(* IEC 61131-3 sources: deprecated-refusr-repo/GP/Main/samples (part 21) *)

(* ---- RND-EXPR_hewed-hoper-pudgy.st ---- *)
(*
This code implements a randomly grown symbolic expression:

((IN43 & IN39) | (!((IN20 & ((IN38 | (!(xor(xor(!(IN25), IN22 | IN24), IN29 | IN3)))) | ((((IN14 | IN14) & (xor(xor(IN1, IN38), IN8))) & (!(IN47 & IN21))) | (IN34 & (xor(xor(xor(xor(IN1, IN18), true), xor(xor(IN14, IN1), IN2)), IN20 | IN27)))))) & ((!(!((xor(xor(!(IN40), !(IN47)), IN24)) | ((IN26 & IN13) | (IN14 | IN31))))) & (!(!(!((!(IN45)) & (!(IN24)))))))))) & ((((xor(xor(IN28, !(IN6)), (xor(xor((xor(xor(true, xor(xor(IN34, IN35), IN30)), IN25 & IN34)) & (IN34 & (!(IN12))), (!(IN38 | IN25)) & IN42), xor(xor(xor(xor(IN20, !(IN31)), IN12), (xor(xor(IN19, IN42), IN21)) & (IN18 & IN20)), (xor(xor(true, IN18), IN13)) & (xor(xor(IN29, IN6), IN10))))) | IN21)) | ((xor(xor(!(((xor(xor(IN4, IN3), IN27)) & IN36) | (IN35 & (!(IN33)))), ((xor(xor(xor(xor(IN12, IN2), IN9), xor(xor(IN39, IN32), IN30)), xor(xor(IN38, IN26), IN25))) | IN26) | (xor(xor((xor(xor(IN37, IN43), IN47)) | IN33, IN1 & (xor(xor(IN11, IN41), IN38))), (IN1 & IN39) | (!(IN13))))), (!(!(!(IN4)))) | (false | ((xor(xor(IN13, IN43), IN36)) | (IN35 | IN32))))) & (IN8 | (!(IN31))))) & (((((xor(xor(xor(xor(IN20, !(IN5)), IN6 | IN30), (IN34 & IN9) | (xor(xor(IN35, IN5), IN16))), xor(xor(IN5, IN3 | IN25), !(IN2)))) & (xor(xor((IN45 | IN10) | (IN49 & IN43), IN20), !(IN2 & IN11)))) | (!((xor(xor(IN17 | IN4, IN25), xor(xor(IN5, IN25), IN16))) & (xor(xor(!(IN43), IN40 & IN25), IN7 | IN48))))) | (IN48 | IN1)) | (!((!((xor(xor(!(IN45), IN8), !(IN21))) | IN34)) | IN9)))) | IN9)

*)

FUNCTION_BLOCK F_CollectInput
  VAR_IN_OUT
      Data : ARRAY[1..50] OF BOOL;
  END_VAR
  VAR_INPUT
      TICK  : BOOL := 0;
      IN1   : BOOL := 0;
      IN2   : BOOL := 0;
      IN3   : BOOL := 0;
      IN4   : BOOL := 0;
      IN5   : BOOL := 0;
      RESET : BOOL := FALSE;
  END_VAR
  VAR_OUTPUT
      Finished : BOOL;
  END_VAR
  VAR
      j    : USINT := 1;
      tock : BOOL  := 0;
  END_VAR
  IF NOT RESET AND tock = NOT TICK THEN
      Data[j]   := IN1;
      Data[j+1] := IN2;
      Data[j+2] := IN3;
      Data[j+3] := IN4;
      Data[j+4] := IN5;
      j := j + 5;
      tock := TICK;
  ELSE
      j := 1;
      tock := 0;
  END_IF;
  Finished := (j > 50);
END_FUNCTION_BLOCK

PROGRAM Boiler
  VAR
    Data  : ARRAY[1..50] OF BOOL;
    Ready : BOOL;
    CollectInput : F_CollectInput;
  END_VAR
  VAR
    TICK     AT %IX1.0 : BOOL;
    IN1      AT %IX0.3 : BOOL;
    IN2      AT %IX0.4 : BOOL;
    IN3      AT %IX0.5 : BOOL;
    IN4      AT %IX0.6 : BOOL;
    IN5      AT %IX0.7 : BOOL;
    OutReady AT %QX0.0 : BOOL := FALSE;
    FeedNext AT %QX0.1 : BOOL := FALSE;
    Out      AT %QX0.2 : BOOL;
  END_VAR
  CollectInput(TICK:=TICK, IN1:=IN1, IN2:=IN2, IN3:=IN3, IN4:=IN4, IN5:=IN5);
  Ready := CollectInput.Finished;
  FeedNext := 1;
  IF Ready THEN
    Out := (((Data[43] AND Data[39]) OR (NOT ((Data[20] AND ((Data[38] OR (NOT (((NOT Data[25]) XOR (Data[22] OR Data[24])) XOR (Data[29] OR Data[3])))) OR ((((Data[14] OR Data[14]) AND ((Data[1] XOR Data[38]) XOR Data[8])) AND (NOT (Data[47] AND Data[21]))) OR (Data[34] AND ((((Data[1] XOR Data[18]) XOR TRUE) XOR ((Data[14] XOR Data[1]) XOR Data[2])) XOR (Data[20] OR Data[27])))))) AND ((NOT (NOT ((((NOT Data[40]) XOR (NOT Data[47])) XOR Data[24]) OR ((Data[26] AND Data[13]) OR (Data[14] OR Data[31]))))) AND (NOT (NOT (NOT ((NOT Data[45]) AND (NOT Data[24]))))))))) AND (((((Data[28] XOR (NOT Data[6])) XOR ((((((TRUE XOR ((Data[34] XOR Data[35]) XOR Data[30])) XOR (Data[25] AND Data[34])) AND (Data[34] AND (NOT Data[12]))) XOR ((NOT (Data[38] OR Data[25])) AND Data[42])) XOR ((((Data[20] XOR (NOT Data[31])) XOR Data[12]) XOR (((Data[19] XOR Data[42]) XOR Data[21]) AND (Data[18] AND Data[20]))) XOR (((TRUE XOR Data[18]) XOR Data[13]) AND ((Data[29] XOR Data[6]) XOR Data[10])))) OR Data[21])) OR ((((NOT ((((Data[4] XOR Data[3]) XOR Data[27]) AND Data[36]) OR (Data[35] AND (NOT Data[33])))) XOR ((((((Data[12] XOR Data[2]) XOR Data[9]) XOR ((Data[39] XOR Data[32]) XOR Data[30])) XOR ((Data[38] XOR Data[26]) XOR Data[25])) OR Data[26]) OR (((((Data[37] XOR Data[43]) XOR Data[47]) OR Data[33]) XOR (Data[1] AND ((Data[11] XOR Data[41]) XOR Data[38]))) XOR ((Data[1] AND Data[39]) OR (NOT Data[13]))))) XOR ((NOT (NOT (NOT Data[4]))) OR (FALSE OR (((Data[13] XOR Data[43]) XOR Data[36]) OR (Data[35] OR Data[32]))))) AND (Data[8] OR (NOT Data[31])))) AND ((((((((Data[20] XOR (NOT Data[5])) XOR (Data[6] OR Data[30])) XOR ((Data[34] AND Data[9]) OR ((Data[35] XOR Data[5]) XOR Data[16]))) XOR ((Data[5] XOR (Data[3] OR Data[25])) XOR (NOT Data[2]))) AND ((((Data[45] OR Data[10]) OR (Data[49] AND Data[43])) XOR Data[20]) XOR (NOT (Data[2] AND Data[11])))) OR (NOT ((((Data[17] OR Data[4]) XOR Data[25]) XOR ((Data[5] XOR Data[25]) XOR Data[16])) AND (((NOT Data[43]) XOR (Data[40] AND Data[25])) XOR (Data[7] OR Data[48]))))) OR (Data[48] OR Data[1])) OR (NOT ((NOT ((((NOT Data[45]) XOR Data[8]) XOR (NOT Data[21])) OR Data[34])) OR Data[9])))) OR Data[9]));
    OutReady := 1;
    CollectInput(RESET:=TRUE);
  END_IF;
END_PROGRAM

CONFIGURATION Config0
  RESOURCE Res0 ON PLC
    TASK task0(INTERVAL := T#20ms,PRIORITY := 0);
    PROGRAM instance0 WITH task0 : Boiler;
  END_RESOURCE
END_CONFIGURATION

(* ---- RND-EXPR_hypos-smote-bongs.st ---- *)
(*
This code implements a randomly grown symbolic expression:

!(((IN8 & (((xor(xor((xor(xor(IN35 & IN19, !(IN2)), IN2)) & ((xor(xor(IN30, IN50), IN41)) | (!(IN35))), ((IN30 & IN28) & (xor(xor(IN2, IN28), IN4))) & (xor(xor(IN18 | IN27, IN9 & IN35), IN12 & IN6))), xor(xor((IN10 & IN14) & (xor(xor(IN6, IN1), IN48)), xor(xor(IN9, IN41 | IN49), false | IN34)), IN31))) & (!(((false | IN35) & IN15) & IN20))) & (xor(xor(IN9, xor(xor(!(IN25), (IN23 & (IN11 | IN39)) | ((IN39 | IN5) | (!(IN26)))), !(!(!(IN38))))), (!(IN1 | (!(IN31)))) | ((IN14 & IN30) & IN6))))) & (!(xor(xor((xor(xor(((!(IN39)) & (true | IN46)) & ((xor(xor(IN13, IN48), IN49)) | (!(IN43))), IN15), !(xor(xor(IN8 & IN6, xor(xor(IN35, IN42), IN13)), IN48 & IN45)))) & (IN17 & (IN26 | (xor(xor(IN39 & false, IN49), !(IN38))))), xor(xor(xor(xor(!(!(!(IN32))), xor(xor(!(xor(xor(IN41, IN2), IN48)), (IN35 & IN6) | (IN29 & IN32)), xor(xor(!(IN22), xor(xor(IN40, IN4), IN36)), IN23 & IN44))), ((IN35 | IN43) | (!(IN38))) | (!(IN26 | IN25))), !((!(IN33 | IN33)) & (xor(xor(xor(xor(IN25, IN3), IN39), IN40), IN26 | IN49)))), IN9)), IN26)))) | ((!((xor(xor(xor(xor(xor(xor((IN27 & IN28) | (IN45 & IN6), (IN25 & IN38) | (IN23 & IN23)), IN48 & (IN40 | IN29)), xor(xor((xor(xor(IN25, IN11), IN33)) & IN36, !(IN40)), xor(xor(IN47 | IN47, !(IN48)), IN30))), IN3), !((IN42 | IN22) & ((IN13 | IN19) & (!(IN22))))), xor(xor(!(IN41 | (IN38 | IN29)), xor(xor(!(IN6 & IN31), IN28), !(xor(xor(IN41, IN32), IN12)))), ((!(IN22)) | (!(IN2))) & (!(IN40 | false))))) | (xor(xor(xor(xor(((IN47 & IN7) & (!(IN19))) & IN3, (!(IN5 & true)) | (!(IN21 & IN16))), ((!(IN12)) & (xor(xor(IN36, IN38), IN43))) & (!(!(IN1)))), IN13), IN11)))) & (!(!((xor(xor(((!(IN5)) & IN1) & IN43, (IN35 & IN17) | IN39), IN32)) & (!(xor(xor(!(!(IN39)), IN13), xor(xor(!(IN20), IN2 & IN50), xor(xor(IN14, IN3), IN25))))))))))

*)

FUNCTION_BLOCK F_CollectInput
  VAR_IN_OUT
      Data : ARRAY[1..50] OF BOOL;
  END_VAR
  VAR_INPUT
      TICK  : BOOL := 0;
      IN1   : BOOL := 0;
      IN2   : BOOL := 0;
      IN3   : BOOL := 0;
      IN4   : BOOL := 0;
      IN5   : BOOL := 0;
      RESET : BOOL := FALSE;
  END_VAR
  VAR_OUTPUT
      Finished : BOOL;
  END_VAR
  VAR
      j    : USINT := 1;
      tock : BOOL  := 0;
  END_VAR
  IF NOT RESET AND tock = NOT TICK THEN
      Data[j]   := IN1;
      Data[j+1] := IN2;
      Data[j+2] := IN3;
      Data[j+3] := IN4;
      Data[j+4] := IN5;
      j := j + 5;
      tock := TICK;
  ELSE
      j := 1;
      tock := 0;
  END_IF;
  Finished := (j > 50);
END_FUNCTION_BLOCK

PROGRAM Boiler
  VAR
    Data  : ARRAY[1..50] OF BOOL;
    Ready : BOOL;
    CollectInput : F_CollectInput;
  END_VAR
  VAR
    TICK     AT %IX1.0 : BOOL;
    IN1      AT %IX0.3 : BOOL;
    IN2      AT %IX0.4 : BOOL;
    IN3      AT %IX0.5 : BOOL;
    IN4      AT %IX0.6 : BOOL;
    IN5      AT %IX0.7 : BOOL;
    OutReady AT %QX0.0 : BOOL := FALSE;
    FeedNext AT %QX0.1 : BOOL := FALSE;
    Out      AT %QX0.2 : BOOL;
  END_VAR
  CollectInput(TICK:=TICK, IN1:=IN1, IN2:=IN2, IN3:=IN3, IN4:=IN4, IN5:=IN5);
  Ready := CollectInput.Finished;
  FeedNext := 1;
  IF Ready THEN
    Out := (NOT (((Data[8] AND ((((((((Data[35] AND Data[19]) XOR (NOT Data[2])) XOR Data[2]) AND (((Data[30] XOR Data[50]) XOR Data[41]) OR (NOT Data[35]))) XOR (((Data[30] AND Data[28]) AND ((Data[2] XOR Data[28]) XOR Data[4])) AND (((Data[18] OR Data[27]) XOR (Data[9] AND Data[35])) XOR (Data[12] AND Data[6])))) XOR ((((Data[10] AND Data[14]) AND ((Data[6] XOR Data[1]) XOR Data[48])) XOR ((Data[9] XOR (Data[41] OR Data[49])) XOR (FALSE OR Data[34]))) XOR Data[31])) AND (NOT (((FALSE OR Data[35]) AND Data[15]) AND Data[20]))) AND ((Data[9] XOR (((NOT Data[25]) XOR ((Data[23] AND (Data[11] OR Data[39])) OR ((Data[39] OR Data[5]) OR (NOT Data[26])))) XOR (NOT (NOT (NOT Data[38]))))) XOR ((NOT (Data[1] OR (NOT Data[31]))) OR ((Data[14] AND Data[30]) AND Data[6]))))) AND (NOT ((((((((NOT Data[39]) AND (TRUE OR Data[46])) AND (((Data[13] XOR Data[48]) XOR Data[49]) OR (NOT Data[43]))) XOR Data[15]) XOR (NOT (((Data[8] AND Data[6]) XOR ((Data[35] XOR Data[42]) XOR Data[13])) XOR (Data[48] AND Data[45])))) AND (Data[17] AND (Data[26] OR (((Data[39] AND FALSE) XOR Data[49]) XOR (NOT Data[38]))))) XOR (((((NOT (NOT (NOT Data[32]))) XOR (((NOT ((Data[41] XOR Data[2]) XOR Data[48])) XOR ((Data[35] AND Data[6]) OR (Data[29] AND Data[32]))) XOR (((NOT Data[22]) XOR ((Data[40] XOR Data[4]) XOR Data[36])) XOR (Data[23] AND Data[44])))) XOR (((Data[35] OR Data[43]) OR (NOT Data[38])) OR (NOT (Data[26] OR Data[25])))) XOR (NOT ((NOT (Data[33] OR Data[33])) AND ((((Data[25] XOR Data[3]) XOR Data[39]) XOR Data[40]) XOR (Data[26] OR Data[49]))))) XOR Data[9])) XOR Data[26]))) OR ((NOT (((((((((Data[27] AND Data[28]) OR (Data[45] AND Data[6])) XOR ((Data[25] AND Data[38]) OR (Data[23] AND Data[23]))) XOR (Data[48] AND (Data[40] OR Data[29]))) XOR (((((Data[25] XOR Data[11]) XOR Data[33]) AND Data[36]) XOR (NOT Data[40])) XOR (((Data[47] OR Data[47]) XOR (NOT Data[48])) XOR Data[30]))) XOR Data[3]) XOR (NOT ((Data[42] OR Data[22]) AND ((Data[13] OR Data[19]) AND (NOT Data[22]))))) XOR (((NOT (Data[41] OR (Data[38] OR Data[29]))) XOR (((NOT (Data[6] AND Data[31])) XOR Data[28]) XOR (NOT ((Data[41] XOR Data[32]) XOR Data[12])))) XOR (((NOT Data[22]) OR (NOT Data[2])) AND (NOT (Data[40] OR FALSE))))) OR (((((((Data[47] AND Data[7]) AND (NOT Data[19])) AND Data[3]) XOR ((NOT (Data[5] AND TRUE)) OR (NOT (Data[21] AND Data[16])))) XOR (((NOT Data[12]) AND ((Data[36] XOR Data[38]) XOR Data[43])) AND (NOT (NOT Data[1])))) XOR Data[13]) XOR Data[11]))) AND (NOT (NOT ((((((NOT Data[5]) AND Data[1]) AND Data[43]) XOR ((Data[35] AND Data[17]) OR Data[39])) XOR Data[32]) AND (NOT (((NOT (NOT Data[39])) XOR Data[13]) XOR (((NOT Data[20]) XOR (Data[2] AND Data[50])) XOR ((Data[14] XOR Data[3]) XOR Data[25]))))))))));
    OutReady := 1;
    CollectInput(RESET:=TRUE);
  END_IF;
END_PROGRAM

CONFIGURATION Config0
  RESOURCE Res0 ON PLC
    TASK task0(INTERVAL := T#20ms,PRIORITY := 0);
    PROGRAM instance0 WITH task0 : Boiler;
  END_RESOURCE
END_CONFIGURATION

(* ---- RND-EXPR_leaky-feued-blurs.st ---- *)
(*
This code implements a randomly grown symbolic expression:

xor(xor(IN1, (xor(xor(xor(xor((!(xor(xor((IN12 | (IN11 & IN27)) & IN11, !(xor(xor(!(IN34), IN44 & IN46), IN19 | IN38))), IN38 | IN45))) | ((IN13 | (xor(xor((xor(xor(IN40, IN15), IN44)) & (IN46 & IN14), IN28 | (xor(xor(IN28, IN38), IN18))), (IN13 & IN4) & (xor(xor(IN22, IN19), IN8))))) | (IN25 & (!((xor(xor(IN10, IN38), IN10)) & (xor(xor(IN42, IN48), IN43)))))), IN21), (IN22 & ((((!(IN41)) | (IN9 & IN29)) & (IN21 & (IN8 & IN45))) | IN6)) & (!(!(!((IN1 & IN39) & IN25))))), (!((xor(xor(IN3 | (false | (!(IN20))), IN30 | ((IN8 & IN45) | (xor(xor(IN44, IN48), IN46)))), (!(!(IN48))) | (!(xor(xor(IN43, IN21), IN14))))) | ((!((IN50 & IN45) | (IN50 | IN41))) | IN42))) & IN39), !(!(xor(xor((IN25 | (xor(xor(IN38, IN38), !(IN48)))) | (((xor(xor(IN26, IN41), true)) & (xor(xor(IN8, IN27), IN34))) | IN15), !(IN40 & (IN44 | (IN13 | IN35)))), IN8))))) & (!(xor(xor(xor(xor((!(IN42)) | (xor(xor((!(IN25 & IN34)) & (xor(xor(IN13 & IN29, IN4 & IN36), !(IN6))), !((IN47 | IN13) & (xor(xor(IN42, IN43), IN40)))), (xor(xor(IN17, IN34), xor(xor(IN8, IN20), IN42))) | ((xor(xor(true, IN21), IN17)) | (!(IN43))))), !(!(((!(IN49)) & (IN44 & IN3)) & (IN20 & (IN6 & IN20))))), !(xor(xor(IN17, IN45), IN32))), ((!(xor(xor((xor(xor(IN4, IN26), IN46)) & (!(IN11)), xor(xor(IN1 | IN28, xor(xor(IN14, IN13), IN41)), !(IN47))), !(IN13)))) | (((xor(xor(!(IN31), IN14 & IN11), xor(xor(IN4, IN7), IN44))) | true) & IN37)) | (xor(xor(!((!(IN40 & IN49)) & IN7), IN15), (IN38 | (xor(xor(IN15, IN33), IN37 | IN17))) & ((xor(xor(IN30 | IN8, IN1), xor(xor(IN9, IN39), IN9))) & ((xor(xor(IN31, IN37), IN48)) & (IN39 | IN29)))))), xor(xor(IN2 | (xor(xor(xor(xor(IN47 & IN29, xor(xor(IN45, IN2), xor(xor(IN47, IN14), IN11))), IN24), !(IN28)), (IN17 | (!(IN48))) | ((xor(xor(IN40, IN45), IN26)) & (IN23 & IN20)))), xor(xor((xor(xor(IN38, !(IN39 | IN3)), IN25 | (xor(xor(IN25, IN3), IN22)))) & (xor(xor((IN2 | true) | (IN39 | IN30), (IN20 & IN40) & (!(IN43))), (IN36 | IN29) | (IN12 | IN39))), !(!(!(!(IN2))))), !(IN41))), (xor(xor(xor(xor((IN5 | IN49) & (!(IN47)), IN19), IN12), IN44), (!(xor(xor(IN23, IN6), IN46))) | (!(IN18 | IN32)))) & (xor(xor((!(!(IN41))) & (IN7 | (false & IN18)), xor(xor(IN49, xor(xor(IN42 | IN42, xor(xor(IN28, IN30), IN31)), xor(xor(IN13, IN37), IN27))), (IN46 | IN24) | (!(IN4)))), (xor(xor(IN33, IN42), !(IN4))) & ((xor(xor(IN24, IN20), IN15)) | (IN22 & IN29))))))))), IN18)

*)

FUNCTION_BLOCK F_CollectInput
  VAR_IN_OUT
      Data : ARRAY[1..50] OF BOOL;
  END_VAR
  VAR_INPUT
      TICK  : BOOL := 0;
      IN1   : BOOL := 0;
      IN2   : BOOL := 0;
      IN3   : BOOL := 0;
      IN4   : BOOL := 0;
      IN5   : BOOL := 0;
      RESET : BOOL := FALSE;
  END_VAR
  VAR_OUTPUT
      Finished : BOOL;
  END_VAR
  VAR
      j    : USINT := 1;
      tock : BOOL  := 0;
  END_VAR
  IF NOT RESET AND tock = NOT TICK THEN
      Data[j]   := IN1;
      Data[j+1] := IN2;
      Data[j+2] := IN3;
      Data[j+3] := IN4;
      Data[j+4] := IN5;
      j := j + 5;
      tock := TICK;
  ELSE
      j := 1;
      tock := 0;
  END_IF;
  Finished := (j > 50);
END_FUNCTION_BLOCK

PROGRAM Boiler
  VAR
    Data  : ARRAY[1..50] OF BOOL;
    Ready : BOOL;
    CollectInput : F_CollectInput;
  END_VAR
  VAR
    TICK     AT %IX1.0 : BOOL;
    IN1      AT %IX0.3 : BOOL;
    IN2      AT %IX0.4 : BOOL;
    IN3      AT %IX0.5 : BOOL;
    IN4      AT %IX0.6 : BOOL;
    IN5      AT %IX0.7 : BOOL;
    OutReady AT %QX0.0 : BOOL := FALSE;
    FeedNext AT %QX0.1 : BOOL := FALSE;
    Out      AT %QX0.2 : BOOL;
  END_VAR
  CollectInput(TICK:=TICK, IN1:=IN1, IN2:=IN2, IN3:=IN3, IN4:=IN4, IN5:=IN5);
  Ready := CollectInput.Finished;
  FeedNext := 1;
  IF Ready THEN
    Out := ((Data[1] XOR (((((((NOT ((((Data[12] OR (Data[11] AND Data[27])) AND Data[11]) XOR (NOT (((NOT Data[34]) XOR (Data[44] AND Data[46])) XOR (Data[19] OR Data[38])))) XOR (Data[38] OR Data[45]))) OR ((Data[13] OR (((((Data[40] XOR Data[15]) XOR Data[44]) AND (Data[46] AND Data[14])) XOR (Data[28] OR ((Data[28] XOR Data[38]) XOR Data[18]))) XOR ((Data[13] AND Data[4]) AND ((Data[22] XOR Data[19]) XOR Data[8])))) OR (Data[25] AND (NOT (((Data[10] XOR Data[38]) XOR Data[10]) AND ((Data[42] XOR Data[48]) XOR Data[43])))))) XOR Data[21]) XOR ((Data[22] AND ((((NOT Data[41]) OR (Data[9] AND Data[29])) AND (Data[21] AND (Data[8] AND Data[45]))) OR Data[6])) AND (NOT (NOT (NOT ((Data[1] AND Data[39]) AND Data[25])))))) XOR ((NOT ((((Data[3] OR (FALSE OR (NOT Data[20]))) XOR (Data[30] OR ((Data[8] AND Data[45]) OR ((Data[44] XOR Data[48]) XOR Data[46])))) XOR ((NOT (NOT Data[48])) OR (NOT ((Data[43] XOR Data[21]) XOR Data[14])))) OR ((NOT ((Data[50] AND Data[45]) OR (Data[50] OR Data[41]))) OR Data[42]))) AND Data[39])) XOR (NOT (NOT ((((Data[25] OR ((Data[38] XOR Data[38]) XOR (NOT Data[48]))) OR ((((Data[26] XOR Data[41]) XOR TRUE) AND ((Data[8] XOR Data[27]) XOR Data[34])) OR Data[15])) XOR (NOT (Data[40] AND (Data[44] OR (Data[13] OR Data[35]))))) XOR Data[8])))) AND (NOT ((((((NOT Data[42]) OR ((((NOT (Data[25] AND Data[34])) AND (((Data[13] AND Data[29]) XOR (Data[4] AND Data[36])) XOR (NOT Data[6]))) XOR (NOT ((Data[47] OR Data[13]) AND ((Data[42] XOR Data[43]) XOR Data[40])))) XOR (((Data[17] XOR Data[34]) XOR ((Data[8] XOR Data[20]) XOR Data[42])) OR (((TRUE XOR Data[21]) XOR Data[17]) OR (NOT Data[43]))))) XOR (NOT (NOT (((NOT Data[49]) AND (Data[44] AND Data[3])) AND (Data[20] AND (Data[6] AND Data[20])))))) XOR (NOT ((Data[17] XOR Data[45]) XOR Data[32]))) XOR (((NOT (((((Data[4] XOR Data[26]) XOR Data[46]) AND (NOT Data[11])) XOR (((Data[1] OR Data[28]) XOR ((Data[14] XOR Data[13]) XOR Data[41])) XOR (NOT Data[47]))) XOR (NOT Data[13]))) OR (((((NOT Data[31]) XOR (Data[14] AND Data[11])) XOR ((Data[4] XOR Data[7]) XOR Data[44])) OR TRUE) AND Data[37])) OR (((NOT ((NOT (Data[40] AND Data[49])) AND Data[7])) XOR Data[15]) XOR ((Data[38] OR ((Data[15] XOR Data[33]) XOR (Data[37] OR Data[17]))) AND ((((Data[30] OR Data[8]) XOR Data[1]) XOR ((Data[9] XOR Data[39]) XOR Data[9])) AND (((Data[31] XOR Data[37]) XOR Data[48]) AND (Data[39] OR Data[29]))))))) XOR (((Data[2] OR (((((Data[47] AND Data[29]) XOR ((Data[45] XOR Data[2]) XOR ((Data[47] XOR Data[14]) XOR Data[11]))) XOR Data[24]) XOR (NOT Data[28])) XOR ((Data[17] OR (NOT Data[48])) OR (((Data[40] XOR Data[45]) XOR Data[26]) AND (Data[23] AND Data[20]))))) XOR (((((Data[38] XOR (NOT (Data[39] OR Data[3]))) XOR (Data[25] OR ((Data[25] XOR Data[3]) XOR Data[22]))) AND ((((Data[2] OR TRUE) OR (Data[39] OR Data[30])) XOR ((Data[20] AND Data[40]) AND (NOT Data[43]))) XOR ((Data[36] OR Data[29]) OR (Data[12] OR Data[39])))) XOR (NOT (NOT (NOT (NOT Data[2]))))) XOR (NOT Data[41]))) XOR (((((((Data[5] OR Data[49]) AND (NOT Data[47])) XOR Data[19]) XOR Data[12]) XOR Data[44]) XOR ((NOT ((Data[23] XOR Data[6]) XOR Data[46])) OR (NOT (Data[18] OR Data[32])))) AND ((((NOT (NOT Data[41])) AND (Data[7] OR (FALSE AND Data[18]))) XOR ((Data[49] XOR (((Data[42] OR Data[42]) XOR ((Data[28] XOR Data[30]) XOR Data[31])) XOR ((Data[13] XOR Data[37]) XOR Data[27]))) XOR ((Data[46] OR Data[24]) OR (NOT Data[4])))) XOR (((Data[33] XOR Data[42]) XOR (NOT Data[4])) AND (((Data[24] XOR Data[20]) XOR Data[15]) OR (Data[22] AND Data[29])))))))))) XOR Data[18]);
    OutReady := 1;
    CollectInput(RESET:=TRUE);
  END_IF;
END_PROGRAM

CONFIGURATION Config0
  RESOURCE Res0 ON PLC
    TASK task0(INTERVAL := T#20ms,PRIORITY := 0);
    PROGRAM instance0 WITH task0 : Boiler;
  END_RESOURCE
END_CONFIGURATION

(* ---- RND-EXPR_limes-bench-plate.st ---- *)
(*
This code implements a randomly grown symbolic expression:

IN28 & (((((xor(xor((!(IN48)) | IN45, ((IN18 | (!(IN46))) | ((!(IN2)) | IN31)) & (xor(xor(!(xor(xor(IN21, IN35), IN5)), !(xor(xor(IN28, false), IN7))), !(IN50 & IN5)))), IN21)) & (((IN1 & ((xor(xor(IN48, IN42), IN3)) & (!(IN22)))) | (xor(xor((!(IN22)) | (xor(xor(IN33, IN36), IN18)), (!(IN25)) & (xor(xor(IN42, IN46), IN34))), !(!(IN3))))) & (xor(xor((!(IN36)) | (!(IN40 | IN41)), IN7), !((!(IN29)) | IN47))))) | ((!(IN3 | ((!(IN1 | IN27)) & (xor(xor(!(IN49), false), !(IN18)))))) | (!(((IN5 | (IN10 & IN32)) & (IN41 | (IN15 | IN22))) | ((xor(xor(xor(xor(IN1, IN10), IN18), !(IN1)), !(IN15))) | ((IN8 & IN5) & (xor(xor(IN1, IN21), IN19)))))))) & (xor(xor(IN36, IN7), ((xor(xor(xor(xor((xor(xor(IN15, IN6), IN17)) & IN2, (IN32 & IN36) & IN19), (xor(xor(false, IN27), IN26)) & (!(IN3))), xor(xor(xor(xor(IN3 & IN45, IN37 & IN38), xor(xor(IN11, IN16), IN32)), (xor(xor(IN48, IN3), IN5)) | IN4), IN29)), IN19)) & (!(xor(xor(IN44, xor(xor(xor(xor(IN36, IN31), IN35), !(IN13)), IN5)), !(IN46 | IN13))))) | IN1))) | (!(!(xor(xor((!(xor(xor(!(IN11 | IN31), !(IN42 | true)), IN42 | (IN42 | IN26)))) | IN7, xor(xor((!(!(IN23 | IN34))) | ((xor(xor(!(IN7), IN5 | IN10), !(IN12))) & ((IN48 | IN15) & (xor(xor(IN31, IN40), IN21)))), (IN24 & (xor(xor(!(IN15), IN26 | IN13), IN38))) | (xor(xor(IN9, (xor(xor(IN39, IN27), IN32)) & (!(IN29))), IN22))), IN30)), IN41)))))

*)

FUNCTION_BLOCK F_CollectInput
  VAR_IN_OUT
      Data : ARRAY[1..50] OF BOOL;
  END_VAR
  VAR_INPUT
      TICK  : BOOL := 0;
      IN1   : BOOL := 0;
      IN2   : BOOL := 0;
      IN3   : BOOL := 0;
      IN4   : BOOL := 0;
      IN5   : BOOL := 0;
      RESET : BOOL := FALSE;
  END_VAR
  VAR_OUTPUT
      Finished : BOOL;
  END_VAR
  VAR
      j    : USINT := 1;
      tock : BOOL  := 0;
  END_VAR
  IF NOT RESET AND tock = NOT TICK THEN
      Data[j]   := IN1;
      Data[j+1] := IN2;
      Data[j+2] := IN3;
      Data[j+3] := IN4;
      Data[j+4] := IN5;
      j := j + 5;
      tock := TICK;
  ELSE
      j := 1;
      tock := 0;
  END_IF;
  Finished := (j > 50);
END_FUNCTION_BLOCK

PROGRAM Boiler
  VAR
    Data  : ARRAY[1..50] OF BOOL;
    Ready : BOOL;
    CollectInput : F_CollectInput;
  END_VAR
  VAR
    TICK     AT %IX1.0 : BOOL;
    IN1      AT %IX0.3 : BOOL;
    IN2      AT %IX0.4 : BOOL;
    IN3      AT %IX0.5 : BOOL;
    IN4      AT %IX0.6 : BOOL;
    IN5      AT %IX0.7 : BOOL;
    OutReady AT %QX0.0 : BOOL := FALSE;
    FeedNext AT %QX0.1 : BOOL := FALSE;
    Out      AT %QX0.2 : BOOL;
  END_VAR
  CollectInput(TICK:=TICK, IN1:=IN1, IN2:=IN2, IN3:=IN3, IN4:=IN4, IN5:=IN5);
  Ready := CollectInput.Finished;
  FeedNext := 1;
  IF Ready THEN
    Out := (Data[28] AND ((((((((NOT Data[48]) OR Data[45]) XOR (((Data[18] OR (NOT Data[46])) OR ((NOT Data[2]) OR Data[31])) AND (((NOT ((Data[21] XOR Data[35]) XOR Data[5])) XOR (NOT ((Data[28] XOR FALSE) XOR Data[7]))) XOR (NOT (Data[50] AND Data[5]))))) XOR Data[21]) AND (((Data[1] AND (((Data[48] XOR Data[42]) XOR Data[3]) AND (NOT Data[22]))) OR ((((NOT Data[22]) OR ((Data[33] XOR Data[36]) XOR Data[18])) XOR ((NOT Data[25]) AND ((Data[42] XOR Data[46]) XOR Data[34]))) XOR (NOT (NOT Data[3])))) AND ((((NOT Data[36]) OR (NOT (Data[40] OR Data[41]))) XOR Data[7]) XOR (NOT ((NOT Data[29]) OR Data[47]))))) OR ((NOT (Data[3] OR ((NOT (Data[1] OR Data[27])) AND (((NOT Data[49]) XOR FALSE) XOR (NOT Data[18]))))) OR (NOT (((Data[5] OR (Data[10] AND Data[32])) AND (Data[41] OR (Data[15] OR Data[22]))) OR (((((Data[1] XOR Data[10]) XOR Data[18]) XOR (NOT Data[1])) XOR (NOT Data[15])) OR ((Data[8] AND Data[5]) AND ((Data[1] XOR Data[21]) XOR Data[19]))))))) AND ((Data[36] XOR Data[7]) XOR (((((((((Data[15] XOR Data[6]) XOR Data[17]) AND Data[2]) XOR ((Data[32] AND Data[36]) AND Data[19])) XOR (((FALSE XOR Data[27]) XOR Data[26]) AND (NOT Data[3]))) XOR (((((Data[3] AND Data[45]) XOR (Data[37] AND Data[38])) XOR ((Data[11] XOR Data[16]) XOR Data[32])) XOR (((Data[48] XOR Data[3]) XOR Data[5]) OR Data[4])) XOR Data[29])) XOR Data[19]) AND (NOT ((Data[44] XOR ((((Data[36] XOR Data[31]) XOR Data[35]) XOR (NOT Data[13])) XOR Data[5])) XOR (NOT (Data[46] OR Data[13]))))) OR Data[1]))) OR (NOT (NOT ((((NOT (((NOT (Data[11] OR Data[31])) XOR (NOT (Data[42] OR TRUE))) XOR (Data[42] OR (Data[42] OR Data[26])))) OR Data[7]) XOR ((((NOT (NOT (Data[23] OR Data[34]))) OR ((((NOT Data[7]) XOR (Data[5] OR Data[10])) XOR (NOT Data[12])) AND ((Data[48] OR Data[15]) AND ((Data[31] XOR Data[40]) XOR Data[21])))) XOR ((Data[24] AND (((NOT Data[15]) XOR (Data[26] OR Data[13])) XOR Data[38])) OR ((Data[9] XOR (((Data[39] XOR Data[27]) XOR Data[32]) AND (NOT Data[29]))) XOR Data[22]))) XOR Data[30])) XOR Data[41])))));
    OutReady := 1;
    CollectInput(RESET:=TRUE);
  END_IF;
END_PROGRAM

CONFIGURATION Config0
  RESOURCE Res0 ON PLC
    TASK task0(INTERVAL := T#20ms,PRIORITY := 0);
    PROGRAM instance0 WITH task0 : Boiler;
  END_RESOURCE
END_CONFIGURATION

(* ---- RND-EXPR_litre-preen-cunts.st ---- *)
(*
This code implements a randomly grown symbolic expression:

!(IN34)

*)

FUNCTION_BLOCK F_CollectInput
  VAR_IN_OUT
      Data : ARRAY[1..50] OF BOOL;
  END_VAR
  VAR_INPUT
      TICK  : BOOL := 0;
      IN1   : BOOL := 0;
      IN2   : BOOL := 0;
      IN3   : BOOL := 0;
      IN4   : BOOL := 0;
      IN5   : BOOL := 0;
      RESET : BOOL := FALSE;
  END_VAR
  VAR_OUTPUT
      Finished : BOOL;
  END_VAR
  VAR
      j    : USINT := 1;
      tock : BOOL  := 0;
  END_VAR
  IF NOT RESET AND tock = NOT TICK THEN
      Data[j]   := IN1;
      Data[j+1] := IN2;
      Data[j+2] := IN3;
      Data[j+3] := IN4;
      Data[j+4] := IN5;
      j := j + 5;
      tock := TICK;
  ELSE
      j := 1;
      tock := 0;
  END_IF;
  Finished := (j > 50);
END_FUNCTION_BLOCK

PROGRAM Boiler
  VAR
    Data  : ARRAY[1..50] OF BOOL;
    Ready : BOOL;
    CollectInput : F_CollectInput;
  END_VAR
  VAR
    TICK     AT %IX1.0 : BOOL;
    IN1      AT %IX0.3 : BOOL;
    IN2      AT %IX0.4 : BOOL;
    IN3      AT %IX0.5 : BOOL;
    IN4      AT %IX0.6 : BOOL;
    IN5      AT %IX0.7 : BOOL;
    OutReady AT %QX0.0 : BOOL := FALSE;
    FeedNext AT %QX0.1 : BOOL := FALSE;
    Out      AT %QX0.2 : BOOL;
  END_VAR
  CollectInput(TICK:=TICK, IN1:=IN1, IN2:=IN2, IN3:=IN3, IN4:=IN4, IN5:=IN5);
  Ready := CollectInput.Finished;
  FeedNext := 1;
  IF Ready THEN
    Out := (NOT Data[34]);
    OutReady := 1;
    CollectInput(RESET:=TRUE);
  END_IF;
END_PROGRAM

CONFIGURATION Config0
  RESOURCE Res0 ON PLC
    TASK task0(INTERVAL := T#20ms,PRIORITY := 0);
    PROGRAM instance0 WITH task0 : Boiler;
  END_RESOURCE
END_CONFIGURATION

(* ---- RND-EXPR_maned-cited-trill.st ---- *)
(*
This code implements a randomly grown symbolic expression:

xor(xor(!(IN14 & (!(!((xor(xor((!(!(IN25))) & ((IN4 | IN27) | IN40), xor(xor(IN45 & IN48, (!(IN36)) | (IN1 & IN33)), !(IN44 | IN43))), IN46 & (xor(xor(IN48 & IN29, IN17 | IN44), IN28 | IN22)))) & ((!((xor(xor(IN22, IN13), IN2)) & (!(IN31)))) | (((IN5 & IN48) & (IN32 & IN20)) & IN29)))))), IN21), xor(xor(xor(xor((xor(xor(!(IN39), (!(!((IN25 | IN46) & (IN25 | IN14)))) | (xor(xor(!(!(!(IN30))), (xor(xor(IN38, !(IN19)), IN16 | IN30)) & IN29), !(!(xor(xor(IN5, IN9), IN17)))))), (!(((xor(xor(IN7, IN10), IN15)) & (xor(xor(IN4, IN7), IN17))) & IN18)) & ((xor(xor(!(IN22 & IN36), (xor(xor(IN49, IN28), IN3)) | IN28), (xor(xor(IN39, IN28), IN36)) | (!(IN29)))) & ((!(IN7 & IN50)) | (!(IN17)))))) | (!(!(IN12))), xor(xor(!((!(IN49)) | (IN2 & IN28)), xor(xor(!((!(IN1)) | IN23), (!(IN2)) & (xor(xor(IN9 & ((IN25 & IN20) | (IN2 & IN27)), IN4), true))), !(((!(xor(xor(IN11, true), IN27))) & (!(IN37 & IN28))) & IN40))), IN11 & IN26)), IN12), xor(xor(IN29, (xor(xor((((xor(xor(IN12 & IN20, !(IN37)), false)) | (!(IN37 & false))) | IN28) | (((xor(xor(IN40 & IN41, IN1), IN37 | IN4)) | ((IN6 | IN48) | (!(IN5)))) & ((xor(xor(!(IN20), !(IN50)), IN37 | IN27)) & (!(!(IN36))))), !(!((xor(xor(!(IN45), !(IN8)), xor(xor(IN35, IN43), IN32))) & ((IN18 & IN14) & (IN17 | IN28))))), (xor(xor(IN50, IN29 | (xor(xor(IN42 | IN32, IN48), IN46 & true))), ((xor(xor(IN8, IN46), IN1)) & (!(IN46))) | (IN49 | IN7))) | (IN2 | ((!(xor(xor(IN8, IN10), IN30))) & (!(xor(xor(IN16, IN30), IN7))))))) & ((((IN4 | ((!(IN38)) | (IN3 | IN19))) | (xor(xor(!(IN46), IN39 & (!(IN35))), xor(xor(xor(xor(IN48, IN12), IN21), !(IN12)), IN41 & IN29)))) | (xor(xor(IN10 | ((!(IN12)) & (IN42 | IN3)), !((IN48 & IN34) | (IN19 | IN22))), xor(xor((!(IN8)) | (IN20 & IN39), IN28 & (IN28 & IN16)), !(xor(xor(IN21, IN12), IN7)))))) | (!(!((IN48 | (!(IN44))) | ((!(IN5)) & (IN49 | IN7))))))), IN2)), !(!((!(xor(xor(((IN13 & IN33) & IN43) | true, (xor(xor(false, IN14 | IN8), IN25 & IN46)) | ((IN46 | IN7) & (IN45 & IN20))), false | ((IN8 & IN27) | (xor(xor(IN24, IN7), IN32)))))) & (xor(xor(xor(xor(IN14, IN39 | (xor(xor(IN37 & IN41, xor(xor(IN39, IN24), IN26)), IN24))), xor(xor(xor(xor(xor(xor(IN49, IN15), IN29), IN7), IN14 & IN13), !(xor(xor(IN28, IN50), IN33))), !(IN27 & IN46))), IN29), (IN13 & IN8) & IN16))))))

*)

FUNCTION_BLOCK F_CollectInput
  VAR_IN_OUT
      Data : ARRAY[1..50] OF BOOL;
  END_VAR
  VAR_INPUT
      TICK  : BOOL := 0;
      IN1   : BOOL := 0;
      IN2   : BOOL := 0;
      IN3   : BOOL := 0;
      IN4   : BOOL := 0;
      IN5   : BOOL := 0;
      RESET : BOOL := FALSE;
  END_VAR
  VAR_OUTPUT
      Finished : BOOL;
  END_VAR
  VAR
      j    : USINT := 1;
      tock : BOOL  := 0;
  END_VAR
  IF NOT RESET AND tock = NOT TICK THEN
      Data[j]   := IN1;
      Data[j+1] := IN2;
      Data[j+2] := IN3;
      Data[j+3] := IN4;
      Data[j+4] := IN5;
      j := j + 5;
      tock := TICK;
  ELSE
      j := 1;
      tock := 0;
  END_IF;
  Finished := (j > 50);
END_FUNCTION_BLOCK

PROGRAM Boiler
  VAR
    Data  : ARRAY[1..50] OF BOOL;
    Ready : BOOL;
    CollectInput : F_CollectInput;
  END_VAR
  VAR
    TICK     AT %IX1.0 : BOOL;
    IN1      AT %IX0.3 : BOOL;
    IN2      AT %IX0.4 : BOOL;
    IN3      AT %IX0.5 : BOOL;
    IN4      AT %IX0.6 : BOOL;
    IN5      AT %IX0.7 : BOOL;
    OutReady AT %QX0.0 : BOOL := FALSE;
    FeedNext AT %QX0.1 : BOOL := FALSE;
    Out      AT %QX0.2 : BOOL;
  END_VAR
  CollectInput(TICK:=TICK, IN1:=IN1, IN2:=IN2, IN3:=IN3, IN4:=IN4, IN5:=IN5);
  Ready := CollectInput.Finished;
  FeedNext := 1;
  IF Ready THEN
    Out := (((NOT (Data[14] AND (NOT (NOT (((((NOT (NOT Data[25])) AND ((Data[4] OR Data[27]) OR Data[40])) XOR (((Data[45] AND Data[48]) XOR ((NOT Data[36]) OR (Data[1] AND Data[33]))) XOR (NOT (Data[44] OR Data[43])))) XOR (Data[46] AND (((Data[48] AND Data[29]) XOR (Data[17] OR Data[44])) XOR (Data[28] OR Data[22])))) AND ((NOT (((Data[22] XOR Data[13]) XOR Data[2]) AND (NOT Data[31]))) OR (((Data[5] AND Data[48]) AND (Data[32] AND Data[20])) AND Data[29]))))))) XOR Data[21]) XOR ((((((((NOT Data[39]) XOR ((NOT (NOT ((Data[25] OR Data[46]) AND (Data[25] OR Data[14])))) OR (((NOT (NOT (NOT Data[30]))) XOR (((Data[38] XOR (NOT Data[19])) XOR (Data[16] OR Data[30])) AND Data[29])) XOR (NOT (NOT ((Data[5] XOR Data[9]) XOR Data[17])))))) XOR ((NOT ((((Data[7] XOR Data[10]) XOR Data[15]) AND ((Data[4] XOR Data[7]) XOR Data[17])) AND Data[18])) AND ((((NOT (Data[22] AND Data[36])) XOR (((Data[49] XOR Data[28]) XOR Data[3]) OR Data[28])) XOR (((Data[39] XOR Data[28]) XOR Data[36]) OR (NOT Data[29]))) AND ((NOT (Data[7] AND Data[50])) OR (NOT Data[17]))))) OR (NOT (NOT Data[12]))) XOR (((NOT ((NOT Data[49]) OR (Data[2] AND Data[28]))) XOR (((NOT ((NOT Data[1]) OR Data[23])) XOR ((NOT Data[2]) AND (((Data[9] AND ((Data[25] AND Data[20]) OR (Data[2] AND Data[27]))) XOR Data[4]) XOR TRUE))) XOR (NOT (((NOT ((Data[11] XOR TRUE) XOR Data[27])) AND (NOT (Data[37] AND Data[28]))) AND Data[40])))) XOR (Data[11] AND Data[26]))) XOR Data[12]) XOR ((Data[29] XOR (((((((((Data[12] AND Data[20]) XOR (NOT Data[37])) XOR FALSE) OR (NOT (Data[37] AND FALSE))) OR Data[28]) OR (((((Data[40] AND Data[41]) XOR Data[1]) XOR (Data[37] OR Data[4])) OR ((Data[6] OR Data[48]) OR (NOT Data[5]))) AND ((((NOT Data[20]) XOR (NOT Data[50])) XOR (Data[37] OR Data[27])) AND (NOT (NOT Data[36]))))) XOR (NOT (NOT ((((NOT Data[45]) XOR (NOT Data[8])) XOR ((Data[35] XOR Data[43]) XOR Data[32])) AND ((Data[18] AND Data[14]) AND (Data[17] OR Data[28])))))) XOR (((Data[50] XOR (Data[29] OR (((Data[42] OR Data[32]) XOR Data[48]) XOR (Data[46] AND TRUE)))) XOR ((((Data[8] XOR Data[46]) XOR Data[1]) AND (NOT Data[46])) OR (Data[49] OR Data[7]))) OR (Data[2] OR ((NOT ((Data[8] XOR Data[10]) XOR Data[30])) AND (NOT ((Data[16] XOR Data[30]) XOR Data[7])))))) AND ((((Data[4] OR ((NOT Data[38]) OR (Data[3] OR Data[19]))) OR (((NOT Data[46]) XOR (Data[39] AND (NOT Data[35]))) XOR ((((Data[48] XOR Data[12]) XOR Data[21]) XOR (NOT Data[12])) XOR (Data[41] AND Data[29])))) OR (((Data[10] OR ((NOT Data[12]) AND (Data[42] OR Data[3]))) XOR (NOT ((Data[48] AND Data[34]) OR (Data[19] OR Data[22])))) XOR ((((NOT Data[8]) OR (Data[20] AND Data[39])) XOR (Data[28] AND (Data[28] AND Data[16]))) XOR (NOT ((Data[21] XOR Data[12]) XOR Data[7]))))) OR (NOT (NOT ((Data[48] OR (NOT Data[44])) OR ((NOT Data[5]) AND (Data[49] OR Data[7])))))))) XOR Data[2])) XOR (NOT (NOT ((NOT (((((Data[13] AND Data[33]) AND Data[43]) OR TRUE) XOR (((FALSE XOR (Data[14] OR Data[8])) XOR (Data[25] AND Data[46])) OR ((Data[46] OR Data[7]) AND (Data[45] AND Data[20])))) XOR (FALSE OR ((Data[8] AND Data[27]) OR ((Data[24] XOR Data[7]) XOR Data[32]))))) AND ((((Data[14] XOR (Data[39] OR (((Data[37] AND Data[41]) XOR ((Data[39] XOR Data[24]) XOR Data[26])) XOR Data[24]))) XOR ((((((Data[49] XOR Data[15]) XOR Data[29]) XOR Data[7]) XOR (Data[14] AND Data[13])) XOR (NOT ((Data[28] XOR Data[50]) XOR Data[33]))) XOR (NOT (Data[27] AND Data[46])))) XOR Data[29]) XOR ((Data[13] AND Data[8]) AND Data[16])))))));
    OutReady := 1;
    CollectInput(RESET:=TRUE);
  END_IF;
END_PROGRAM

CONFIGURATION Config0
  RESOURCE Res0 ON PLC
    TASK task0(INTERVAL := T#20ms,PRIORITY := 0);
    PROGRAM instance0 WITH task0 : Boiler;
  END_RESOURCE
END_CONFIGURATION

(* ---- RND-EXPR_mason-gases-tombs.st ---- *)
(*
This code implements a randomly grown symbolic expression:

((!(xor(xor(xor(xor(IN36, (!((!(xor(xor(IN22, IN23), IN42))) & (!(IN43 & IN13)))) & IN27), IN22), !(!((xor(xor(xor(xor(xor(xor(IN41, IN40), IN6), IN18 | IN25), xor(xor(IN48, IN48), IN11)), !(IN30 & IN33)), (!(IN46)) | (xor(xor(IN33, IN43), IN34)))) | (((IN2 | IN35) & (IN31 & IN45)) & ((IN24 & IN42) | (IN23 & IN28)))))), (IN14 | IN11) & (xor(xor((!(IN19)) & (!((IN6 & IN28) | IN32)), (!(!(IN33 | IN45))) & (((xor(xor(IN46, IN13), IN17)) & (!(IN24))) | (!(IN36 | IN10)))), xor(xor(IN11, IN45 | ((xor(xor(IN34, IN31), IN18)) & (!(IN24)))), !(!(!(IN48))))))))) | (xor(xor(xor(xor(xor(xor(IN27, IN7), IN45), IN36), IN7 | ((xor(xor(((IN17 & IN37) | (IN41 | IN20)) & (!(xor(xor(IN28, IN28), IN43))), IN41 & ((IN50 | IN20) | (IN16 & IN43))), (xor(xor(IN30, IN46), IN5 & IN10)) & ((!(IN22)) & (xor(xor(IN9, true), IN2))))) | (!(xor(xor(xor(xor(!(IN44), !(IN39)), !(IN14)), (!(IN21)) | (!(IN50))), xor(xor(xor(xor(IN6, IN4), IN36), IN25 & IN10), !(IN34))))))), IN29), (!(IN30)) & IN6))) & IN10

*)

FUNCTION_BLOCK F_CollectInput
  VAR_IN_OUT
      Data : ARRAY[1..50] OF BOOL;
  END_VAR
  VAR_INPUT
      TICK  : BOOL := 0;
      IN1   : BOOL := 0;
      IN2   : BOOL := 0;
      IN3   : BOOL := 0;
      IN4   : BOOL := 0;
      IN5   : BOOL := 0;
      RESET : BOOL := FALSE;
  END_VAR
  VAR_OUTPUT
      Finished : BOOL;
  END_VAR
  VAR
      j    : USINT := 1;
      tock : BOOL  := 0;
  END_VAR
  IF NOT RESET AND tock = NOT TICK THEN
      Data[j]   := IN1;
      Data[j+1] := IN2;
      Data[j+2] := IN3;
      Data[j+3] := IN4;
      Data[j+4] := IN5;
      j := j + 5;
      tock := TICK;
  ELSE
      j := 1;
      tock := 0;
  END_IF;
  Finished := (j > 50);
END_FUNCTION_BLOCK

PROGRAM Boiler
  VAR
    Data  : ARRAY[1..50] OF BOOL;
    Ready : BOOL;
    CollectInput : F_CollectInput;
  END_VAR
  VAR
    TICK     AT %IX1.0 : BOOL;
    IN1      AT %IX0.3 : BOOL;
    IN2      AT %IX0.4 : BOOL;
    IN3      AT %IX0.5 : BOOL;
    IN4      AT %IX0.6 : BOOL;
    IN5      AT %IX0.7 : BOOL;
    OutReady AT %QX0.0 : BOOL := FALSE;
    FeedNext AT %QX0.1 : BOOL := FALSE;
    Out      AT %QX0.2 : BOOL;
  END_VAR
  CollectInput(TICK:=TICK, IN1:=IN1, IN2:=IN2, IN3:=IN3, IN4:=IN4, IN5:=IN5);
  Ready := CollectInput.Finished;
  FeedNext := 1;
  IF Ready THEN
    Out := (((NOT ((((Data[36] XOR ((NOT ((NOT ((Data[22] XOR Data[23]) XOR Data[42])) AND (NOT (Data[43] AND Data[13])))) AND Data[27])) XOR Data[22]) XOR (NOT (NOT (((((((Data[41] XOR Data[40]) XOR Data[6]) XOR (Data[18] OR Data[25])) XOR ((Data[48] XOR Data[48]) XOR Data[11])) XOR (NOT (Data[30] AND Data[33]))) XOR ((NOT Data[46]) OR ((Data[33] XOR Data[43]) XOR Data[34]))) OR (((Data[2] OR Data[35]) AND (Data[31] AND Data[45])) AND ((Data[24] AND Data[42]) OR (Data[23] AND Data[28]))))))) XOR ((Data[14] OR Data[11]) AND ((((NOT Data[19]) AND (NOT ((Data[6] AND Data[28]) OR Data[32]))) XOR ((NOT (NOT (Data[33] OR Data[45]))) AND ((((Data[46] XOR Data[13]) XOR Data[17]) AND (NOT Data[24])) OR (NOT (Data[36] OR Data[10]))))) XOR ((Data[11] XOR (Data[45] OR (((Data[34] XOR Data[31]) XOR Data[18]) AND (NOT Data[24])))) XOR (NOT (NOT (NOT Data[48])))))))) OR ((((((Data[27] XOR Data[7]) XOR Data[45]) XOR Data[36]) XOR (Data[7] OR ((((((Data[17] AND Data[37]) OR (Data[41] OR Data[20])) AND (NOT ((Data[28] XOR Data[28]) XOR Data[43]))) XOR (Data[41] AND ((Data[50] OR Data[20]) OR (Data[16] AND Data[43])))) XOR (((Data[30] XOR Data[46]) XOR (Data[5] AND Data[10])) AND ((NOT Data[22]) AND ((Data[9] XOR TRUE) XOR Data[2])))) OR (NOT (((((NOT Data[44]) XOR (NOT Data[39])) XOR (NOT Data[14])) XOR ((NOT Data[21]) OR (NOT Data[50]))) XOR ((((Data[6] XOR Data[4]) XOR Data[36]) XOR (Data[25] AND Data[10])) XOR (NOT Data[34]))))))) XOR Data[29]) XOR ((NOT Data[30]) AND Data[6]))) AND Data[10]);
    OutReady := 1;
    CollectInput(RESET:=TRUE);
  END_IF;
END_PROGRAM

CONFIGURATION Config0
  RESOURCE Res0 ON PLC
    TASK task0(INTERVAL := T#20ms,PRIORITY := 0);
    PROGRAM instance0 WITH task0 : Boiler;
  END_RESOURCE
END_CONFIGURATION

(* ---- RND-EXPR_maven-hello-baize.st ---- *)
(*
This code implements a randomly grown symbolic expression:

((!(!(IN21 & (xor(xor(false, !(!((xor(xor(false, IN2), IN25)) | (!(IN9))))), ((IN33 & (xor(xor(IN17, IN40), IN11))) & (xor(xor(xor(xor(IN20, IN38), IN8), IN28 & IN33), IN19 & IN13))) & IN13))))) & IN25) & ((!((xor(xor(IN28, xor(xor((!(!(IN8 | IN21))) | ((!(IN47 | IN48)) | (!(IN15))), (!(IN9)) | ((xor(xor(IN49 & IN47, IN49 & IN24), IN46 | IN22)) | (!(IN28)))), !(((IN34 & IN44) & IN48) & IN26))), !(xor(xor(!((xor(xor(IN22, IN48), IN19)) | IN13), IN46), !((xor(xor(IN22, IN42), IN14)) | IN16))))) & ((((xor(xor((false | IN22) & (IN6 & IN36), (!(IN36)) & (IN1 & IN42)), IN21 & IN2)) | IN42) | IN48) | (!(IN36))))) & (IN15 | ((xor(xor(!(!(xor(xor((IN30 | IN11) | (IN43 & IN31), IN43 & (IN50 | IN12)), (IN13 & IN46) | (IN47 & IN18)))), ((IN47 | ((!(IN45)) & IN30)) & (xor(xor(xor(xor(IN6, IN1 & IN6), IN47), xor(xor(IN1 | IN29, IN33), false)), IN35))) | (xor(xor(((!(IN21)) | (!(IN25))) & (IN46 & (IN9 | IN19)), xor(xor(!(IN12 | IN11), xor(xor(IN8 & IN17, IN35 & IN20), xor(xor(IN38, IN14), IN18))), IN36 | (IN49 | IN43))), xor(xor((IN5 & IN20) & (xor(xor(IN20, IN17), IN15)), (xor(xor(IN2, IN24), IN37)) & IN6), IN18 & (IN41 | IN4))))), !(xor(xor(IN3, IN35), (xor(xor(IN29 & IN48, xor(xor(IN41, IN30), IN24)), IN15 | IN43)) | ((!(IN29)) | (false | IN42)))))) & (!(!(IN21 | (((!(IN38)) | (IN48 | IN49)) | IN16)))))))

*)

FUNCTION_BLOCK F_CollectInput
  VAR_IN_OUT
      Data : ARRAY[1..50] OF BOOL;
  END_VAR
  VAR_INPUT
      TICK  : BOOL := 0;
      IN1   : BOOL := 0;
      IN2   : BOOL := 0;
      IN3   : BOOL := 0;
      IN4   : BOOL := 0;
      IN5   : BOOL := 0;
      RESET : BOOL := FALSE;
  END_VAR
  VAR_OUTPUT
      Finished : BOOL;
  END_VAR
  VAR
      j    : USINT := 1;
      tock : BOOL  := 0;
  END_VAR
  IF NOT RESET AND tock = NOT TICK THEN
      Data[j]   := IN1;
      Data[j+1] := IN2;
      Data[j+2] := IN3;
      Data[j+3] := IN4;
      Data[j+4] := IN5;
      j := j + 5;
      tock := TICK;
  ELSE
      j := 1;
      tock := 0;
  END_IF;
  Finished := (j > 50);
END_FUNCTION_BLOCK

PROGRAM Boiler
  VAR
    Data  : ARRAY[1..50] OF BOOL;
    Ready : BOOL;
    CollectInput : F_CollectInput;
  END_VAR
  VAR
    TICK     AT %IX1.0 : BOOL;
    IN1      AT %IX0.3 : BOOL;
    IN2      AT %IX0.4 : BOOL;
    IN3      AT %IX0.5 : BOOL;
    IN4      AT %IX0.6 : BOOL;
    IN5      AT %IX0.7 : BOOL;
    OutReady AT %QX0.0 : BOOL := FALSE;
    FeedNext AT %QX0.1 : BOOL := FALSE;
    Out      AT %QX0.2 : BOOL;
  END_VAR
  CollectInput(TICK:=TICK, IN1:=IN1, IN2:=IN2, IN3:=IN3, IN4:=IN4, IN5:=IN5);
  Ready := CollectInput.Finished;
  FeedNext := 1;
  IF Ready THEN
    Out := (((NOT (NOT (Data[21] AND ((FALSE XOR (NOT (NOT (((FALSE XOR Data[2]) XOR Data[25]) OR (NOT Data[9]))))) XOR (((Data[33] AND ((Data[17] XOR Data[40]) XOR Data[11])) AND ((((Data[20] XOR Data[38]) XOR Data[8]) XOR (Data[28] AND Data[33])) XOR (Data[19] AND Data[13]))) AND Data[13]))))) AND Data[25]) AND ((NOT (((Data[28] XOR ((((NOT (NOT (Data[8] OR Data[21]))) OR ((NOT (Data[47] OR Data[48])) OR (NOT Data[15]))) XOR ((NOT Data[9]) OR ((((Data[49] AND Data[47]) XOR (Data[49] AND Data[24])) XOR (Data[46] OR Data[22])) OR (NOT Data[28])))) XOR (NOT (((Data[34] AND Data[44]) AND Data[48]) AND Data[26])))) XOR (NOT (((NOT (((Data[22] XOR Data[48]) XOR Data[19]) OR Data[13])) XOR Data[46]) XOR (NOT (((Data[22] XOR Data[42]) XOR Data[14]) OR Data[16]))))) AND (((((((FALSE OR Data[22]) AND (Data[6] AND Data[36])) XOR ((NOT Data[36]) AND (Data[1] AND Data[42]))) XOR (Data[21] AND Data[2])) OR Data[42]) OR Data[48]) OR (NOT Data[36])))) AND (Data[15] OR ((((NOT (NOT ((((Data[30] OR Data[11]) OR (Data[43] AND Data[31])) XOR (Data[43] AND (Data[50] OR Data[12]))) XOR ((Data[13] AND Data[46]) OR (Data[47] AND Data[18]))))) XOR (((Data[47] OR ((NOT Data[45]) AND Data[30])) AND ((((Data[6] XOR (Data[1] AND Data[6])) XOR Data[47]) XOR (((Data[1] OR Data[29]) XOR Data[33]) XOR FALSE)) XOR Data[35])) OR (((((NOT Data[21]) OR (NOT Data[25])) AND (Data[46] AND (Data[9] OR Data[19]))) XOR (((NOT (Data[12] OR Data[11])) XOR (((Data[8] AND Data[17]) XOR (Data[35] AND Data[20])) XOR ((Data[38] XOR Data[14]) XOR Data[18]))) XOR (Data[36] OR (Data[49] OR Data[43])))) XOR ((((Data[5] AND Data[20]) AND ((Data[20] XOR Data[17]) XOR Data[15])) XOR (((Data[2] XOR Data[24]) XOR Data[37]) AND Data[6])) XOR (Data[18] AND (Data[41] OR Data[4])))))) XOR (NOT ((Data[3] XOR Data[35]) XOR ((((Data[29] AND Data[48]) XOR ((Data[41] XOR Data[30]) XOR Data[24])) XOR (Data[15] OR Data[43])) OR ((NOT Data[29]) OR (FALSE OR Data[42])))))) AND (NOT (NOT (Data[21] OR (((NOT Data[38]) OR (Data[48] OR Data[49])) OR Data[16]))))))));
    OutReady := 1;
    CollectInput(RESET:=TRUE);
  END_IF;
END_PROGRAM

CONFIGURATION Config0
  RESOURCE Res0 ON PLC
    TASK task0(INTERVAL := T#20ms,PRIORITY := 0);
    PROGRAM instance0 WITH task0 : Boiler;
  END_RESOURCE
END_CONFIGURATION

(* ---- RND-EXPR_mavis-chows-pagan.st ---- *)
(*
This code implements a randomly grown symbolic expression:

!(((xor(xor(((!((xor(xor(IN5 & IN31, IN14), xor(xor(IN41, IN34), IN36))) | (xor(xor(IN5 & true, xor(xor(IN20, IN11), IN46)), xor(xor(IN9, IN25), IN28))))) | ((!((IN16 | IN46) | (IN34 | IN14))) & (((!(IN2)) & (IN5 | IN10)) | (xor(xor(xor(xor(IN46, IN24), IN5), IN28), xor(xor(IN22, IN7), IN13)))))) | (!(IN19 | (xor(xor((!(IN12)) | (IN2 & IN50), IN16), (IN45 & IN28) & IN21)))), xor(xor((xor(xor((xor(xor(IN6 & IN27, IN43 | IN5), IN28)) | (!(IN20 | IN22)), (IN35 & (IN50 | IN10)) | (!(IN19 & IN2))), IN7)) & (!(xor(xor((IN40 | IN16) & (xor(xor(IN27, IN8), IN19)), (xor(xor(IN45, IN13), IN13)) | (IN25 | IN3)), xor(xor(!(IN49), IN29 & IN12), IN16)))), ((!(xor(xor(xor(xor(IN33, IN26), IN50), !(IN42)), !(IN30)))) & IN3) & (xor(xor(!(xor(xor(IN2, xor(xor(false, IN16), true)), xor(xor(IN17, IN11), IN10))), IN24), ((IN41 | IN26) & (!(IN44))) & (!(!(IN6)))))), IN30 & IN4)), xor(xor(xor(xor(!((xor(xor(xor(xor(IN31, IN12), IN9), IN26 | IN38), xor(xor(IN20, IN24), IN46))) | ((IN20 & true) & IN13)), (!(IN36)) | (xor(xor(xor(xor(xor(xor(IN2, IN48), IN8), xor(xor(IN24, IN16), IN9)), IN50 & IN17), IN49), (xor(xor(IN31, true), IN31)) | (xor(xor(IN16, IN38), IN3))))), IN32), IN39), xor(xor((IN17 & (xor(xor(IN35, IN17), !(IN22)))) & (!((!(IN41)) | (IN28 | true))), xor(xor(((!(IN13)) & (xor(xor(IN29, IN36), IN8))) | (xor(xor(IN23 | IN37, IN18 | IN30), IN14 & IN24)), IN39), IN35)), (((IN5 | IN5) & (xor(xor(IN38, IN9), IN45))) & (xor(xor(xor(xor(IN14, IN9), IN1), xor(xor(IN3, IN7), IN34)), !(IN5)))) & ((xor(xor(true | IN3, IN49), IN17 | IN7)) | (!(xor(xor(IN29, IN5), IN48)))))))) | ((xor(xor(xor(xor(xor(xor(!((xor(xor(IN22, IN48), IN22)) | (xor(xor(IN2, true), IN15))), !(IN23)), false), !(((!(IN29)) | (IN46 & IN10)) & ((IN43 | IN35) & IN45))), IN5), (((!(IN35 & true)) | IN22) | (IN39 & (xor(xor(!(IN23), !(IN14)), IN5)))) | (false & (((true & IN42) | (xor(xor(IN16, IN12), IN19))) & (xor(xor(IN5 | IN16, !(IN31)), IN13 & IN46))))), xor(xor(((xor(xor(false & IN31, !(IN12)), IN38)) | ((IN12 & IN14) & IN26)) | (IN14 & (xor(xor(IN42 | IN16, IN50 | IN20), IN1 | IN31))), ((xor(xor(IN44 & IN16, IN29 & IN26), IN19)) & (xor(xor(IN17 & IN46, !(IN42)), xor(xor(IN40, IN42), IN9)))) & ((xor(xor(IN16, !(IN41)), IN2 & IN40)) | ((IN36 | IN3) | IN49))), ((xor(xor(IN35 & IN9, IN19 & IN34), IN12 | IN47)) & ((IN45 & IN19) & (!(IN33)))) | (((IN40 | IN32) | (IN2 | true)) & (xor(xor(IN40 & IN15, xor(xor(IN30, IN5), IN35)), IN48 & IN16)))))) & (!((xor(xor(IN16, IN15), !(!(true & IN45)))) & ((((!(IN44)) | (IN16 & IN26)) | IN43) | (((xor(xor(IN42, IN39), IN40)) | (IN42 & IN8)) & (xor(xor(IN37 & IN7, !(IN1)), IN30 | IN24)))))))) | (!(IN24)))

*)

FUNCTION_BLOCK F_CollectInput
  VAR_IN_OUT
      Data : ARRAY[1..50] OF BOOL;
  END_VAR
  VAR_INPUT
      TICK  : BOOL := 0;
      IN1   : BOOL := 0;
      IN2   : BOOL := 0;
      IN3   : BOOL := 0;
      IN4   : BOOL := 0;
      IN5   : BOOL := 0;
      RESET : BOOL := FALSE;
  END_VAR
  VAR_OUTPUT
      Finished : BOOL;
  END_VAR
  VAR
      j    : USINT := 1;
      tock : BOOL  := 0;
  END_VAR
  IF NOT RESET AND tock = NOT TICK THEN
      Data[j]   := IN1;
      Data[j+1] := IN2;
      Data[j+2] := IN3;
      Data[j+3] := IN4;
      Data[j+4] := IN5;
      j := j + 5;
      tock := TICK;
  ELSE
      j := 1;
      tock := 0;
  END_IF;
  Finished := (j > 50);
END_FUNCTION_BLOCK

PROGRAM Boiler
  VAR
    Data  : ARRAY[1..50] OF BOOL;
    Ready : BOOL;
    CollectInput : F_CollectInput;
  END_VAR
  VAR
    TICK     AT %IX1.0 : BOOL;
    IN1      AT %IX0.3 : BOOL;
    IN2      AT %IX0.4 : BOOL;
    IN3      AT %IX0.5 : BOOL;
    IN4      AT %IX0.6 : BOOL;
    IN5      AT %IX0.7 : BOOL;
    OutReady AT %QX0.0 : BOOL := FALSE;
    FeedNext AT %QX0.1 : BOOL := FALSE;
    Out      AT %QX0.2 : BOOL;
  END_VAR
  CollectInput(TICK:=TICK, IN1:=IN1, IN2:=IN2, IN3:=IN3, IN4:=IN4, IN5:=IN5);
  Ready := CollectInput.Finished;
  FeedNext := 1;
  IF Ready THEN
    Out := (NOT (((((((NOT ((((Data[5] AND Data[31]) XOR Data[14]) XOR ((Data[41] XOR Data[34]) XOR Data[36])) OR (((Data[5] AND TRUE) XOR ((Data[20] XOR Data[11]) XOR Data[46])) XOR ((Data[9] XOR Data[25]) XOR Data[28])))) OR ((NOT ((Data[16] OR Data[46]) OR (Data[34] OR Data[14]))) AND (((NOT Data[2]) AND (Data[5] OR Data[10])) OR ((((Data[46] XOR Data[24]) XOR Data[5]) XOR Data[28]) XOR ((Data[22] XOR Data[7]) XOR Data[13]))))) OR (NOT (Data[19] OR ((((NOT Data[12]) OR (Data[2] AND Data[50])) XOR Data[16]) XOR ((Data[45] AND Data[28]) AND Data[21]))))) XOR (((((((((Data[6] AND Data[27]) XOR (Data[43] OR Data[5])) XOR Data[28]) OR (NOT (Data[20] OR Data[22]))) XOR ((Data[35] AND (Data[50] OR Data[10])) OR (NOT (Data[19] AND Data[2])))) XOR Data[7]) AND (NOT ((((Data[40] OR Data[16]) AND ((Data[27] XOR Data[8]) XOR Data[19])) XOR (((Data[45] XOR Data[13]) XOR Data[13]) OR (Data[25] OR Data[3]))) XOR (((NOT Data[49]) XOR (Data[29] AND Data[12])) XOR Data[16])))) XOR (((NOT ((((Data[33] XOR Data[26]) XOR Data[50]) XOR (NOT Data[42])) XOR (NOT Data[30]))) AND Data[3]) AND (((NOT ((Data[2] XOR ((FALSE XOR Data[16]) XOR TRUE)) XOR ((Data[17] XOR Data[11]) XOR Data[10]))) XOR Data[24]) XOR (((Data[41] OR Data[26]) AND (NOT Data[44])) AND (NOT (NOT Data[6])))))) XOR (Data[30] AND Data[4]))) XOR (((((NOT (((((Data[31] XOR Data[12]) XOR Data[9]) XOR (Data[26] OR Data[38])) XOR ((Data[20] XOR Data[24]) XOR Data[46])) OR ((Data[20] AND TRUE) AND Data[13]))) XOR ((NOT Data[36]) OR ((((((Data[2] XOR Data[48]) XOR Data[8]) XOR ((Data[24] XOR Data[16]) XOR Data[9])) XOR (Data[50] AND Data[17])) XOR Data[49]) XOR (((Data[31] XOR TRUE) XOR Data[31]) OR ((Data[16] XOR Data[38]) XOR Data[3]))))) XOR Data[32]) XOR Data[39]) XOR ((((Data[17] AND ((Data[35] XOR Data[17]) XOR (NOT Data[22]))) AND (NOT ((NOT Data[41]) OR (Data[28] OR TRUE)))) XOR (((((NOT Data[13]) AND ((Data[29] XOR Data[36]) XOR Data[8])) OR (((Data[23] OR Data[37]) XOR (Data[18] OR Data[30])) XOR (Data[14] AND Data[24]))) XOR Data[39]) XOR Data[35])) XOR ((((Data[5] OR Data[5]) AND ((Data[38] XOR Data[9]) XOR Data[45])) AND ((((Data[14] XOR Data[9]) XOR Data[1]) XOR ((Data[3] XOR Data[7]) XOR Data[34])) XOR (NOT Data[5]))) AND ((((TRUE OR Data[3]) XOR Data[49]) XOR (Data[17] OR Data[7])) OR (NOT ((Data[29] XOR Data[5]) XOR Data[48]))))))) OR ((((((((NOT (((Data[22] XOR Data[48]) XOR Data[22]) OR ((Data[2] XOR TRUE) XOR Data[15]))) XOR (NOT Data[23])) XOR FALSE) XOR (NOT (((NOT Data[29]) OR (Data[46] AND Data[10])) AND ((Data[43] OR Data[35]) AND Data[45])))) XOR Data[5]) XOR ((((NOT (Data[35] AND TRUE)) OR Data[22]) OR (Data[39] AND (((NOT Data[23]) XOR (NOT Data[14])) XOR Data[5]))) OR (FALSE AND (((TRUE AND Data[42]) OR ((Data[16] XOR Data[12]) XOR Data[19])) AND (((Data[5] OR Data[16]) XOR (NOT Data[31])) XOR (Data[13] AND Data[46])))))) XOR (((((((FALSE AND Data[31]) XOR (NOT Data[12])) XOR Data[38]) OR ((Data[12] AND Data[14]) AND Data[26])) OR (Data[14] AND (((Data[42] OR Data[16]) XOR (Data[50] OR Data[20])) XOR (Data[1] OR Data[31])))) XOR (((((Data[44] AND Data[16]) XOR (Data[29] AND Data[26])) XOR Data[19]) AND (((Data[17] AND Data[46]) XOR (NOT Data[42])) XOR ((Data[40] XOR Data[42]) XOR Data[9]))) AND (((Data[16] XOR (NOT Data[41])) XOR (Data[2] AND Data[40])) OR ((Data[36] OR Data[3]) OR Data[49])))) XOR (((((Data[35] AND Data[9]) XOR (Data[19] AND Data[34])) XOR (Data[12] OR Data[47])) AND ((Data[45] AND Data[19]) AND (NOT Data[33]))) OR (((Data[40] OR Data[32]) OR (Data[2] OR TRUE)) AND (((Data[40] AND Data[15]) XOR ((Data[30] XOR Data[5]) XOR Data[35])) XOR (Data[48] AND Data[16])))))) AND (NOT (((Data[16] XOR Data[15]) XOR (NOT (NOT (TRUE AND Data[45])))) AND ((((NOT Data[44]) OR (Data[16] AND Data[26])) OR Data[43]) OR ((((Data[42] XOR Data[39]) XOR Data[40]) OR (Data[42] AND Data[8])) AND (((Data[37] AND Data[7]) XOR (NOT Data[1])) XOR (Data[30] OR Data[24])))))))) OR (NOT Data[24])));
    OutReady := 1;
    CollectInput(RESET:=TRUE);
  END_IF;
END_PROGRAM

CONFIGURATION Config0
  RESOURCE Res0 ON PLC
    TASK task0(INTERVAL := T#20ms,PRIORITY := 0);
    PROGRAM instance0 WITH task0 : Boiler;
  END_RESOURCE
END_CONFIGURATION

(* ---- RND-EXPR_medal-trams-sprig.st ---- *)
(*
This code implements a randomly grown symbolic expression:

(!(IN9 & IN6)) | ((xor(xor(IN42, xor(xor(xor(xor((((xor(xor(IN21 & IN3, !(IN48)), IN25)) & ((IN25 | IN29) & (!(IN34)))) & (!(xor(xor(!(IN8), IN43 | IN34), true & IN3)))) & (IN30 & IN22), true), xor(xor(IN11, IN23), !(IN20))), !(xor(xor(xor(xor((!(IN23 | IN23)) & ((IN7 | IN35) | (xor(xor(IN10, IN11), IN30))), !((IN48 | IN22) | (IN18 & IN41))), !((!(IN24)) & (xor(xor(IN11, IN46), IN30)))), IN3), (xor(xor((IN10 | IN30) & (xor(xor(IN44, IN23), IN34)), (xor(xor(IN49, IN33), IN38)) | (IN23 | IN38)), IN20)) | ((xor(xor(xor(xor(IN34, IN10), IN39), xor(xor(IN18, IN42), IN17)), IN17 | IN30)) | IN44)))), (!(IN36)) & (((xor(xor(xor(xor(IN38 | IN4, IN48 | IN16), IN48), (xor(xor(IN24, IN18), false)) & IN14), (xor(xor(IN35, IN22), IN4)) | (IN6 | IN42))) | IN6) | (xor(xor(!(!(IN47)), (xor(xor(IN25 & IN33, !(IN19)), !(IN43))) | ((IN3 & IN6) | true)), xor(xor(IN44, (IN40 | IN1) & (!(IN46))), IN25)))))), xor(xor((xor(xor(IN14, xor(xor(IN3, (xor(xor(!(IN35), xor(xor(IN29, IN2), IN25)), xor(xor(IN43, IN27), IN1))) & ((IN32 | IN35) & IN17)), true & ((IN45 & IN30) & IN39))), (((xor(xor(IN7, IN43), IN40)) & (IN43 | IN5)) | (!(IN13 | IN2))) & (((!(IN47)) & (IN49 | IN50)) | (IN38 | (!(IN48)))))) & (xor(xor(xor(xor(IN24 | ((!(IN23)) | (IN11 & IN7)), ((IN37 & IN42) | (IN5 | IN11)) | ((IN46 & IN36) | (IN27 & IN27))), xor(xor((IN33 & IN37) & (!(IN46)), IN48 & (IN38 & IN49)), (xor(xor(IN15, IN17), IN33)) | (IN25 | IN34))), !(((xor(xor(IN46, IN21), IN11)) | (xor(xor(IN8, IN34), false))) & (xor(xor(xor(xor(false, IN1), IN37), xor(xor(false, IN23), IN23)), IN44)))), !(((IN39 & IN12) & (xor(xor(IN48, IN2), IN22))) | (xor(xor(IN16, true), !(IN19)))))), (((((IN38 | IN31) & (xor(xor(IN39, IN8), IN24))) | ((IN35 & IN18) | (IN34 & IN3))) | ((xor(xor(IN34 | IN30, xor(xor(IN41, IN33), IN25)), IN36 | IN31)) | ((false & IN29) & (!(IN8))))) & IN10) & (xor(xor(IN16, xor(xor(((IN13 & IN2) | (IN5 & IN25)) | (xor(xor(IN41 | IN38, IN38 | true), !(IN18))), (!(IN30 | IN15)) & (!(IN30 | IN24))), xor(xor(IN3, xor(xor(xor(xor(IN34, IN19), IN22), xor(xor(IN35, IN16), IN26)), !(IN10))), (IN49 & IN6) | (IN49 | IN10)))), IN47))), (((!((!(IN30)) & IN4)) | (!(!(IN42 | IN10)))) | IN50) | (IN11 & ((xor(xor(IN8, (!(IN6)) & (IN1 | IN42)), !(xor(xor(IN9, IN23), IN10)))) | (!((IN26 & IN21) & IN32))))))) | (!(!((!(IN23)) & (((((IN15 | IN15) | (IN14 & false)) & (xor(xor(xor(xor(IN34, IN16), IN27), IN10 & IN45), xor(xor(IN45, IN30), IN11)))) | (IN10 | ((IN7 | IN3) | IN30))) | (xor(xor(xor(xor(xor(xor(IN37, IN41 | IN7), IN44 | IN10), IN8), xor(xor(xor(xor(IN50, IN34), IN27), xor(xor(IN39, IN44), IN36)), xor(xor(IN16, IN37), IN18))), IN47), ((xor(xor(IN10, IN38), IN24)) | (IN22 | IN25)) | (xor(xor(IN41, IN17), IN1 & IN50)))))))))

*)

FUNCTION_BLOCK F_CollectInput
  VAR_IN_OUT
      Data : ARRAY[1..50] OF BOOL;
  END_VAR
  VAR_INPUT
      TICK  : BOOL := 0;
      IN1   : BOOL := 0;
      IN2   : BOOL := 0;
      IN3   : BOOL := 0;
      IN4   : BOOL := 0;
      IN5   : BOOL := 0;
      RESET : BOOL := FALSE;
  END_VAR
  VAR_OUTPUT
      Finished : BOOL;
  END_VAR
  VAR
      j    : USINT := 1;
      tock : BOOL  := 0;
  END_VAR
  IF NOT RESET AND tock = NOT TICK THEN
      Data[j]   := IN1;
      Data[j+1] := IN2;
      Data[j+2] := IN3;
      Data[j+3] := IN4;
      Data[j+4] := IN5;
      j := j + 5;
      tock := TICK;
  ELSE
      j := 1;
      tock := 0;
  END_IF;
  Finished := (j > 50);
END_FUNCTION_BLOCK

PROGRAM Boiler
  VAR
    Data  : ARRAY[1..50] OF BOOL;
    Ready : BOOL;
    CollectInput : F_CollectInput;
  END_VAR
  VAR
    TICK     AT %IX1.0 : BOOL;
    IN1      AT %IX0.3 : BOOL;
    IN2      AT %IX0.4 : BOOL;
    IN3      AT %IX0.5 : BOOL;
    IN4      AT %IX0.6 : BOOL;
    IN5      AT %IX0.7 : BOOL;
    OutReady AT %QX0.0 : BOOL := FALSE;
    FeedNext AT %QX0.1 : BOOL := FALSE;
    Out      AT %QX0.2 : BOOL;
  END_VAR
  CollectInput(TICK:=TICK, IN1:=IN1, IN2:=IN2, IN3:=IN3, IN4:=IN4, IN5:=IN5);
  Ready := CollectInput.Finished;
  FeedNext := 1;
  IF Ready THEN
    Out := ((NOT (Data[9] AND Data[6])) OR (((Data[42] XOR ((((((((((Data[21] AND Data[3]) XOR (NOT Data[48])) XOR Data[25]) AND ((Data[25] OR Data[29]) AND (NOT Data[34]))) AND (NOT (((NOT Data[8]) XOR (Data[43] OR Data[34])) XOR (TRUE AND Data[3])))) AND (Data[30] AND Data[22])) XOR TRUE) XOR ((Data[11] XOR Data[23]) XOR (NOT Data[20]))) XOR (NOT ((((((NOT (Data[23] OR Data[23])) AND ((Data[7] OR Data[35]) OR ((Data[10] XOR Data[11]) XOR Data[30]))) XOR (NOT ((Data[48] OR Data[22]) OR (Data[18] AND Data[41])))) XOR (NOT ((NOT Data[24]) AND ((Data[11] XOR Data[46]) XOR Data[30])))) XOR Data[3]) XOR (((((Data[10] OR Data[30]) AND ((Data[44] XOR Data[23]) XOR Data[34])) XOR (((Data[49] XOR Data[33]) XOR Data[38]) OR (Data[23] OR Data[38]))) XOR Data[20]) OR (((((Data[34] XOR Data[10]) XOR Data[39]) XOR ((Data[18] XOR Data[42]) XOR Data[17])) XOR (Data[17] OR Data[30])) OR Data[44]))))) XOR ((NOT Data[36]) AND (((((((Data[38] OR Data[4]) XOR (Data[48] OR Data[16])) XOR Data[48]) XOR (((Data[24] XOR Data[18]) XOR FALSE) AND Data[14])) XOR (((Data[35] XOR Data[22]) XOR Data[4]) OR (Data[6] OR Data[42]))) OR Data[6]) OR (((NOT (NOT Data[47])) XOR ((((Data[25] AND Data[33]) XOR (NOT Data[19])) XOR (NOT Data[43])) OR ((Data[3] AND Data[6]) OR TRUE))) XOR ((Data[44] XOR ((Data[40] OR Data[1]) AND (NOT Data[46]))) XOR Data[25])))))) XOR (((((Data[14] XOR ((Data[3] XOR ((((NOT Data[35]) XOR ((Data[29] XOR Data[2]) XOR Data[25])) XOR ((Data[43] XOR Data[27]) XOR Data[1])) AND ((Data[32] OR Data[35]) AND Data[17]))) XOR (TRUE AND ((Data[45] AND Data[30]) AND Data[39])))) XOR (((((Data[7] XOR Data[43]) XOR Data[40]) AND (Data[43] OR Data[5])) OR (NOT (Data[13] OR Data[2]))) AND (((NOT Data[47]) AND (Data[49] OR Data[50])) OR (Data[38] OR (NOT Data[48]))))) AND (((((Data[24] OR ((NOT Data[23]) OR (Data[11] AND Data[7]))) XOR (((Data[37] AND Data[42]) OR (Data[5] OR Data[11])) OR ((Data[46] AND Data[36]) OR (Data[27] AND Data[27])))) XOR ((((Data[33] AND Data[37]) AND (NOT Data[46])) XOR (Data[48] AND (Data[38] AND Data[49]))) XOR (((Data[15] XOR Data[17]) XOR Data[33]) OR (Data[25] OR Data[34])))) XOR (NOT ((((Data[46] XOR Data[21]) XOR Data[11]) OR ((Data[8] XOR Data[34]) XOR FALSE)) AND ((((FALSE XOR Data[1]) XOR Data[37]) XOR ((FALSE XOR Data[23]) XOR Data[23])) XOR Data[44])))) XOR (NOT (((Data[39] AND Data[12]) AND ((Data[48] XOR Data[2]) XOR Data[22])) OR ((Data[16] XOR TRUE) XOR (NOT Data[19])))))) XOR ((((((Data[38] OR Data[31]) AND ((Data[39] XOR Data[8]) XOR Data[24])) OR ((Data[35] AND Data[18]) OR (Data[34] AND Data[3]))) OR ((((Data[34] OR Data[30]) XOR ((Data[41] XOR Data[33]) XOR Data[25])) XOR (Data[36] OR Data[31])) OR ((FALSE AND Data[29]) AND (NOT Data[8])))) AND Data[10]) AND ((Data[16] XOR (((((Data[13] AND Data[2]) OR (Data[5] AND Data[25])) OR (((Data[41] OR Data[38]) XOR (Data[38] OR TRUE)) XOR (NOT Data[18]))) XOR ((NOT (Data[30] OR Data[15])) AND (NOT (Data[30] OR Data[24])))) XOR ((Data[3] XOR ((((Data[34] XOR Data[19]) XOR Data[22]) XOR ((Data[35] XOR Data[16]) XOR Data[26])) XOR (NOT Data[10]))) XOR ((Data[49] AND Data[6]) OR (Data[49] OR Data[10]))))) XOR Data[47]))) XOR ((((NOT ((NOT Data[30]) AND Data[4])) OR (NOT (NOT (Data[42] OR Data[10])))) OR Data[50]) OR (Data[11] AND (((Data[8] XOR ((NOT Data[6]) AND (Data[1] OR Data[42]))) XOR (NOT ((Data[9] XOR Data[23]) XOR Data[10]))) OR (NOT ((Data[26] AND Data[21]) AND Data[32]))))))) OR (NOT (NOT ((NOT Data[23]) AND (((((Data[15] OR Data[15]) OR (Data[14] AND FALSE)) AND ((((Data[34] XOR Data[16]) XOR Data[27]) XOR (Data[10] AND Data[45])) XOR ((Data[45] XOR Data[30]) XOR Data[11]))) OR (Data[10] OR ((Data[7] OR Data[3]) OR Data[30]))) OR ((((((Data[37] XOR (Data[41] OR Data[7])) XOR (Data[44] OR Data[10])) XOR Data[8]) XOR ((((Data[50] XOR Data[34]) XOR Data[27]) XOR ((Data[39] XOR Data[44]) XOR Data[36])) XOR ((Data[16] XOR Data[37]) XOR Data[18]))) XOR Data[47]) XOR ((((Data[10] XOR Data[38]) XOR Data[24]) OR (Data[22] OR Data[25])) OR ((Data[41] XOR Data[17]) XOR (Data[1] AND Data[50]))))))))));
    OutReady := 1;
    CollectInput(RESET:=TRUE);
  END_IF;
END_PROGRAM

CONFIGURATION Config0
  RESOURCE Res0 ON PLC
    TASK task0(INTERVAL := T#20ms,PRIORITY := 0);
    PROGRAM instance0 WITH task0 : Boiler;
  END_RESOURCE
END_CONFIGURATION

(* ---- RND-EXPR_midst-gauze-lacer.st ---- *)
(*
This code implements a randomly grown symbolic expression:

(!(xor(xor(xor(xor(IN4, IN14), IN32 & ((xor(xor(true, IN23), ((!(IN31)) & (IN21 & IN2)) & IN4)) | IN15)), ((!((xor(xor(IN10, !(IN22 | false)), (xor(xor(IN19, false), IN39)) | (xor(xor(IN50, IN43), IN25)))) | (xor(xor((IN43 | IN12) & (IN48 | IN12), (false & IN12) & IN36), xor(xor(xor(xor(IN8, IN14), IN49), xor(xor(IN10, IN6), IN8)), IN40 & false))))) & (IN23 | ((((IN13 & IN26) | (!(IN33))) | ((!(IN41)) | (IN5 | IN16))) & (!(!(IN32 & IN47)))))) | ((IN24 & (!(!((!(IN20)) | (xor(xor(IN18, IN25), IN29)))))) & IN36)), xor(xor(!(IN39), (((xor(xor(xor(xor(IN11 | IN50, xor(xor(IN49, IN22), IN6)), !(IN21)), !(IN26 | IN40)), (!(IN40)) | IN15)) | (!((IN42 & IN6) & IN14))) & (IN19 & (((IN11 | IN42) | (!(IN36))) & ((IN31 & IN38) & (IN4 & IN20))))) | (((xor(xor((IN39 | IN6) & IN28, (IN43 | IN26) & (IN20 & IN5)), IN25 & (!(IN7)))) | IN34) & ((xor(xor(IN44, !(IN42 | IN15)), xor(xor(IN13 & IN35, IN38 & IN49), IN3 & IN47))) | (!(IN32))))), (!((!(IN45 | (xor(xor(IN25, IN17), IN7)))) | (!((xor(xor(IN6, IN12), IN22)) | (IN27 & IN49))))) & IN20)))) | ((!(IN6)) | (xor(xor((((xor(xor(((xor(xor(IN20, IN3), IN24)) & (!(IN29))) & (xor(xor(IN48 & IN19, xor(xor(IN39, IN26), IN12)), IN20 | IN33)), (IN29 & (xor(xor(IN21, IN47), IN10))) & (!(xor(xor(IN23, IN10), IN45)))), ((!(IN5)) | (!(IN35))) | (!(IN17 | IN44)))) | IN18) | (IN21 & (!(IN4 & IN41)))) & IN42, xor(xor((xor(xor(!(((xor(xor(IN4, IN15), IN42)) | (IN8 | IN5)) | (!(IN25 | IN47))), ((!(xor(xor(IN49, IN22), IN5))) & (xor(xor(IN48, !(IN44)), IN8))) | ((xor(xor(IN24 | IN31, IN42 & IN43), xor(xor(IN47, IN50), IN41))) & (IN25 & (IN20 & IN48)))), xor(xor(((true | IN6) & (!(IN30))) | ((xor(xor(IN15, IN30), IN12)) & (true | IN37)), IN3), xor(xor(xor(xor(false, IN32 & IN50), IN17 | IN37), (IN27 & IN27) & (IN18 | IN25)), IN40 | (IN12 & IN33))))) | (((IN36 & ((IN1 & IN8) | (IN17 | IN48))) | (!(xor(xor(IN32 & IN41, xor(xor(IN28, IN7), IN46)), IN14)))) | IN3), !(((xor(xor(xor(xor(!(IN9), IN40 & IN45), IN33), !(IN39)), IN43)) | ((xor(xor(IN48, IN34 | IN14), IN49 & IN3)) & (IN24 | (IN2 & true)))) | ((xor(xor(IN47, !(IN38)), !(IN13 | IN17))) | (!((xor(xor(IN20, IN32), IN40)) | (!(IN19))))))), (((IN22 | ((IN31 | IN11) & (xor(xor(IN35, false), IN47)))) & (((!(IN22)) & (xor(xor(IN2, IN33), IN45))) & (xor(xor(xor(xor(true, IN46), IN10), IN14 & IN41), IN5 & IN8)))) | (xor(xor(!(IN45), xor(xor(IN49, xor(xor(!(IN36), xor(xor(IN9, IN23), IN26)), IN29 & IN47)), (xor(xor(IN30, IN40), IN49)) & (IN15 & IN42))), (!(IN22 | IN25)) | ((!(IN8)) | (!(IN42)))))) & IN39)), (IN8 | (((((!(IN5)) & (IN44 & IN27)) | ((!(IN43)) | (IN42 & IN17))) & ((xor(xor(IN20 & IN46, IN36), !(IN6))) | ((xor(xor(IN45, false), IN40)) | (!(IN24))))) | (!(((IN13 | IN49) | (true & IN16)) & IN3)))) & ((!(!((!(IN16 & IN1)) | (xor(xor(IN33, xor(xor(IN6, IN28), IN2)), xor(xor(IN31, IN19), IN26)))))) & (IN40 | false)))))

*)

FUNCTION_BLOCK F_CollectInput
  VAR_IN_OUT
      Data : ARRAY[1..50] OF BOOL;
  END_VAR
  VAR_INPUT
      TICK  : BOOL := 0;
      IN1   : BOOL := 0;
      IN2   : BOOL := 0;
      IN3   : BOOL := 0;
      IN4   : BOOL := 0;
      IN5   : BOOL := 0;
      RESET : BOOL := FALSE;
  END_VAR
  VAR_OUTPUT
      Finished : BOOL;
  END_VAR
  VAR
      j    : USINT := 1;
      tock : BOOL  := 0;
  END_VAR
  IF NOT RESET AND tock = NOT TICK THEN
      Data[j]   := IN1;
      Data[j+1] := IN2;
      Data[j+2] := IN3;
      Data[j+3] := IN4;
      Data[j+4] := IN5;
      j := j + 5;
      tock := TICK;
  ELSE
      j := 1;
      tock := 0;
  END_IF;
  Finished := (j > 50);
END_FUNCTION_BLOCK

PROGRAM Boiler
  VAR
    Data  : ARRAY[1..50] OF BOOL;
    Ready : BOOL;
    CollectInput : F_CollectInput;
  END_VAR
  VAR
    TICK     AT %IX1.0 : BOOL;
    IN1      AT %IX0.3 : BOOL;
    IN2      AT %IX0.4 : BOOL;
    IN3      AT %IX0.5 : BOOL;
    IN4      AT %IX0.6 : BOOL;
    IN5      AT %IX0.7 : BOOL;
    OutReady AT %QX0.0 : BOOL := FALSE;
    FeedNext AT %QX0.1 : BOOL := FALSE;
    Out      AT %QX0.2 : BOOL;
  END_VAR
  CollectInput(TICK:=TICK, IN1:=IN1, IN2:=IN2, IN3:=IN3, IN4:=IN4, IN5:=IN5);
  Ready := CollectInput.Finished;
  FeedNext := 1;
  IF Ready THEN
    Out := ((NOT ((((Data[4] XOR Data[14]) XOR (Data[32] AND (((TRUE XOR Data[23]) XOR (((NOT Data[31]) AND (Data[21] AND Data[2])) AND Data[4])) OR Data[15]))) XOR (((NOT (((Data[10] XOR (NOT (Data[22] OR FALSE))) XOR (((Data[19] XOR FALSE) XOR Data[39]) OR ((Data[50] XOR Data[43]) XOR Data[25]))) OR ((((Data[43] OR Data[12]) AND (Data[48] OR Data[12])) XOR ((FALSE AND Data[12]) AND Data[36])) XOR ((((Data[8] XOR Data[14]) XOR Data[49]) XOR ((Data[10] XOR Data[6]) XOR Data[8])) XOR (Data[40] AND FALSE))))) AND (Data[23] OR ((((Data[13] AND Data[26]) OR (NOT Data[33])) OR ((NOT Data[41]) OR (Data[5] OR Data[16]))) AND (NOT (NOT (Data[32] AND Data[47])))))) OR ((Data[24] AND (NOT (NOT ((NOT Data[20]) OR ((Data[18] XOR Data[25]) XOR Data[29]))))) AND Data[36]))) XOR (((NOT Data[39]) XOR ((((((((Data[11] OR Data[50]) XOR ((Data[49] XOR Data[22]) XOR Data[6])) XOR (NOT Data[21])) XOR (NOT (Data[26] OR Data[40]))) XOR ((NOT Data[40]) OR Data[15])) OR (NOT ((Data[42] AND Data[6]) AND Data[14]))) AND (Data[19] AND (((Data[11] OR Data[42]) OR (NOT Data[36])) AND ((Data[31] AND Data[38]) AND (Data[4] AND Data[20]))))) OR ((((((Data[39] OR Data[6]) AND Data[28]) XOR ((Data[43] OR Data[26]) AND (Data[20] AND Data[5]))) XOR (Data[25] AND (NOT Data[7]))) OR Data[34]) AND (((Data[44] XOR (NOT (Data[42] OR Data[15]))) XOR (((Data[13] AND Data[35]) XOR (Data[38] AND Data[49])) XOR (Data[3] AND Data[47]))) OR (NOT Data[32]))))) XOR ((NOT ((NOT (Data[45] OR ((Data[25] XOR Data[17]) XOR Data[7]))) OR (NOT (((Data[6] XOR Data[12]) XOR Data[22]) OR (Data[27] AND Data[49]))))) AND Data[20])))) OR ((NOT Data[6]) OR (((((((((((Data[20] XOR Data[3]) XOR Data[24]) AND (NOT Data[29])) AND (((Data[48] AND Data[19]) XOR ((Data[39] XOR Data[26]) XOR Data[12])) XOR (Data[20] OR Data[33]))) XOR ((Data[29] AND ((Data[21] XOR Data[47]) XOR Data[10])) AND (NOT ((Data[23] XOR Data[10]) XOR Data[45])))) XOR (((NOT Data[5]) OR (NOT Data[35])) OR (NOT (Data[17] OR Data[44])))) OR Data[18]) OR (Data[21] AND (NOT (Data[4] AND Data[41])))) AND Data[42]) XOR ((((((NOT ((((Data[4] XOR Data[15]) XOR Data[42]) OR (Data[8] OR Data[5])) OR (NOT (Data[25] OR Data[47])))) XOR (((NOT ((Data[49] XOR Data[22]) XOR Data[5])) AND ((Data[48] XOR (NOT Data[44])) XOR Data[8])) OR ((((Data[24] OR Data[31]) XOR (Data[42] AND Data[43])) XOR ((Data[47] XOR Data[50]) XOR Data[41])) AND (Data[25] AND (Data[20] AND Data[48]))))) XOR (((((TRUE OR Data[6]) AND (NOT Data[30])) OR (((Data[15] XOR Data[30]) XOR Data[12]) AND (TRUE OR Data[37]))) XOR Data[3]) XOR ((((FALSE XOR (Data[32] AND Data[50])) XOR (Data[17] OR Data[37])) XOR ((Data[27] AND Data[27]) AND (Data[18] OR Data[25]))) XOR (Data[40] OR (Data[12] AND Data[33]))))) OR (((Data[36] AND ((Data[1] AND Data[8]) OR (Data[17] OR Data[48]))) OR (NOT (((Data[32] AND Data[41]) XOR ((Data[28] XOR Data[7]) XOR Data[46])) XOR Data[14]))) OR Data[3])) XOR (NOT (((((((NOT Data[9]) XOR (Data[40] AND Data[45])) XOR Data[33]) XOR (NOT Data[39])) XOR Data[43]) OR (((Data[48] XOR (Data[34] OR Data[14])) XOR (Data[49] AND Data[3])) AND (Data[24] OR (Data[2] AND TRUE)))) OR (((Data[47] XOR (NOT Data[38])) XOR (NOT (Data[13] OR Data[17]))) OR (NOT (((Data[20] XOR Data[32]) XOR Data[40]) OR (NOT Data[19]))))))) XOR ((((Data[22] OR ((Data[31] OR Data[11]) AND ((Data[35] XOR FALSE) XOR Data[47]))) AND (((NOT Data[22]) AND ((Data[2] XOR Data[33]) XOR Data[45])) AND ((((TRUE XOR Data[46]) XOR Data[10]) XOR (Data[14] AND Data[41])) XOR (Data[5] AND Data[8])))) OR (((NOT Data[45]) XOR ((Data[49] XOR (((NOT Data[36]) XOR ((Data[9] XOR Data[23]) XOR Data[26])) XOR (Data[29] AND Data[47]))) XOR (((Data[30] XOR Data[40]) XOR Data[49]) AND (Data[15] AND Data[42])))) XOR ((NOT (Data[22] OR Data[25])) OR ((NOT Data[8]) OR (NOT Data[42]))))) AND Data[39]))) XOR ((Data[8] OR (((((NOT Data[5]) AND (Data[44] AND Data[27])) OR ((NOT Data[43]) OR (Data[42] AND Data[17]))) AND ((((Data[20] AND Data[46]) XOR Data[36]) XOR (NOT Data[6])) OR (((Data[45] XOR FALSE) XOR Data[40]) OR (NOT Data[24])))) OR (NOT (((Data[13] OR Data[49]) OR (TRUE AND Data[16])) AND Data[3])))) AND ((NOT (NOT ((NOT (Data[16] AND Data[1])) OR ((Data[33] XOR ((Data[6] XOR Data[28]) XOR Data[2])) XOR ((Data[31] XOR Data[19]) XOR Data[26]))))) AND (Data[40] OR FALSE))))));
    OutReady := 1;
    CollectInput(RESET:=TRUE);
  END_IF;
END_PROGRAM

CONFIGURATION Config0
  RESOURCE Res0 ON PLC
    TASK task0(INTERVAL := T#20ms,PRIORITY := 0);
    PROGRAM instance0 WITH task0 : Boiler;
  END_RESOURCE
END_CONFIGURATION

(* ---- RND-EXPR_midst-recap-stern.st ---- *)
(*
This code implements a randomly grown symbolic expression:

!(IN41)

*)

FUNCTION_BLOCK F_CollectInput
  VAR_IN_OUT
      Data : ARRAY[1..50] OF BOOL;
  END_VAR
  VAR_INPUT
      TICK  : BOOL := 0;
      IN1   : BOOL := 0;
      IN2   : BOOL := 0;
      IN3   : BOOL := 0;
      IN4   : BOOL := 0;
      IN5   : BOOL := 0;
      RESET : BOOL := FALSE;
  END_VAR
  VAR_OUTPUT
      Finished : BOOL;
  END_VAR
  VAR
      j    : USINT := 1;
      tock : BOOL  := 0;
  END_VAR
  IF NOT RESET AND tock = NOT TICK THEN
      Data[j]   := IN1;
      Data[j+1] := IN2;
      Data[j+2] := IN3;
      Data[j+3] := IN4;
      Data[j+4] := IN5;
      j := j + 5;
      tock := TICK;
  ELSE
      j := 1;
      tock := 0;
  END_IF;
  Finished := (j > 50);
END_FUNCTION_BLOCK

PROGRAM Boiler
  VAR
    Data  : ARRAY[1..50] OF BOOL;
    Ready : BOOL;
    CollectInput : F_CollectInput;
  END_VAR
  VAR
    TICK     AT %IX1.0 : BOOL;
    IN1      AT %IX0.3 : BOOL;
    IN2      AT %IX0.4 : BOOL;
    IN3      AT %IX0.5 : BOOL;
    IN4      AT %IX0.6 : BOOL;
    IN5      AT %IX0.7 : BOOL;
    OutReady AT %QX0.0 : BOOL := FALSE;
    FeedNext AT %QX0.1 : BOOL := FALSE;
    Out      AT %QX0.2 : BOOL;
  END_VAR
  CollectInput(TICK:=TICK, IN1:=IN1, IN2:=IN2, IN3:=IN3, IN4:=IN4, IN5:=IN5);
  Ready := CollectInput.Finished;
  FeedNext := 1;
  IF Ready THEN
    Out := (NOT Data[41]);
    OutReady := 1;
    CollectInput(RESET:=TRUE);
  END_IF;
END_PROGRAM

CONFIGURATION Config0
  RESOURCE Res0 ON PLC
    TASK task0(INTERVAL := T#20ms,PRIORITY := 0);
    PROGRAM instance0 WITH task0 : Boiler;
  END_RESOURCE
END_CONFIGURATION

(* ---- RND-EXPR_mires-marsh-cured.st ---- *)
(*
This code implements a randomly grown symbolic expression:

!(((!(xor(xor(IN30, (xor(xor((xor(xor(IN16 | IN8, IN8), xor(xor(IN24, IN38), IN7))) & (xor(xor(!(IN21), IN44 & IN20), IN50 & IN12)), xor(xor((xor(xor(IN35, IN2), IN16)) | IN3, (IN35 & IN44) | (!(IN2))), !(IN37 & IN50))), !(xor(xor(IN23, false), !(IN16))))) | (xor(xor(IN36, (!(IN10 | IN3)) | ((!(IN48)) & (!(IN25)))), xor(xor(!(IN37 & IN4), (IN25 | IN36) & IN11), IN5 & (IN38 & IN39))))), !(!(!(xor(xor(xor(xor(IN18, IN39), IN11), IN12 | IN44), IN27 | IN37))))))) & (!((!(xor(xor(IN15 | ((xor(xor(IN42, IN3), IN46)) | (xor(xor(IN47, IN27), IN37))), xor(xor(IN1, (IN29 | IN42) & IN43), IN26)), IN21))) | (xor(xor(IN39, ((IN19 | (xor(xor(IN18, IN35), IN2))) | (IN7 & (!(IN24)))) | ((xor(xor(xor(xor(IN44, true), IN45), IN32 & IN47), IN38 & IN43)) & (!(IN40 | IN47)))), xor(xor((!(IN37)) & ((!(IN32)) | (!(IN50))), IN24), !(!(IN42)))))))) | IN5)

*)

FUNCTION_BLOCK F_CollectInput
  VAR_IN_OUT
      Data : ARRAY[1..50] OF BOOL;
  END_VAR
  VAR_INPUT
      TICK  : BOOL := 0;
      IN1   : BOOL := 0;
      IN2   : BOOL := 0;
      IN3   : BOOL := 0;
      IN4   : BOOL := 0;
      IN5   : BOOL := 0;
      RESET : BOOL := FALSE;
  END_VAR
  VAR_OUTPUT
      Finished : BOOL;
  END_VAR
  VAR
      j    : USINT := 1;
      tock : BOOL  := 0;
  END_VAR
  IF NOT RESET AND tock = NOT TICK THEN
      Data[j]   := IN1;
      Data[j+1] := IN2;
      Data[j+2] := IN3;
      Data[j+3] := IN4;
      Data[j+4] := IN5;
      j := j + 5;
      tock := TICK;
  ELSE
      j := 1;
      tock := 0;
  END_IF;
  Finished := (j > 50);
END_FUNCTION_BLOCK

PROGRAM Boiler
  VAR
    Data  : ARRAY[1..50] OF BOOL;
    Ready : BOOL;
    CollectInput : F_CollectInput;
  END_VAR
  VAR
    TICK     AT %IX1.0 : BOOL;
    IN1      AT %IX0.3 : BOOL;
    IN2      AT %IX0.4 : BOOL;
    IN3      AT %IX0.5 : BOOL;
    IN4      AT %IX0.6 : BOOL;
    IN5      AT %IX0.7 : BOOL;
    OutReady AT %QX0.0 : BOOL := FALSE;
    FeedNext AT %QX0.1 : BOOL := FALSE;
    Out      AT %QX0.2 : BOOL;
  END_VAR
  CollectInput(TICK:=TICK, IN1:=IN1, IN2:=IN2, IN3:=IN3, IN4:=IN4, IN5:=IN5);
  Ready := CollectInput.Finished;
  FeedNext := 1;
  IF Ready THEN
    Out := (NOT (((NOT ((Data[30] XOR (((((((Data[16] OR Data[8]) XOR Data[8]) XOR ((Data[24] XOR Data[38]) XOR Data[7])) AND (((NOT Data[21]) XOR (Data[44] AND Data[20])) XOR (Data[50] AND Data[12]))) XOR (((((Data[35] XOR Data[2]) XOR Data[16]) OR Data[3]) XOR ((Data[35] AND Data[44]) OR (NOT Data[2]))) XOR (NOT (Data[37] AND Data[50])))) XOR (NOT ((Data[23] XOR FALSE) XOR (NOT Data[16])))) OR ((Data[36] XOR ((NOT (Data[10] OR Data[3])) OR ((NOT Data[48]) AND (NOT Data[25])))) XOR (((NOT (Data[37] AND Data[4])) XOR ((Data[25] OR Data[36]) AND Data[11])) XOR (Data[5] AND (Data[38] AND Data[39])))))) XOR (NOT (NOT (NOT ((((Data[18] XOR Data[39]) XOR Data[11]) XOR (Data[12] OR Data[44])) XOR (Data[27] OR Data[37]))))))) AND (NOT ((NOT (((Data[15] OR (((Data[42] XOR Data[3]) XOR Data[46]) OR ((Data[47] XOR Data[27]) XOR Data[37]))) XOR ((Data[1] XOR ((Data[29] OR Data[42]) AND Data[43])) XOR Data[26])) XOR Data[21])) OR ((Data[39] XOR (((Data[19] OR ((Data[18] XOR Data[35]) XOR Data[2])) OR (Data[7] AND (NOT Data[24]))) OR (((((Data[44] XOR TRUE) XOR Data[45]) XOR (Data[32] AND Data[47])) XOR (Data[38] AND Data[43])) AND (NOT (Data[40] OR Data[47]))))) XOR ((((NOT Data[37]) AND ((NOT Data[32]) OR (NOT Data[50]))) XOR Data[24]) XOR (NOT (NOT Data[42]))))))) OR Data[5]));
    OutReady := 1;
    CollectInput(RESET:=TRUE);
  END_IF;
END_PROGRAM

CONFIGURATION Config0
  RESOURCE Res0 ON PLC
    TASK task0(INTERVAL := T#20ms,PRIORITY := 0);
    PROGRAM instance0 WITH task0 : Boiler;
  END_RESOURCE
END_CONFIGURATION

(* ---- RND-EXPR_mitre-whews-wraps.st ---- *)
(*
This code implements a randomly grown symbolic expression:

!(!(IN11 | IN43))

*)

FUNCTION_BLOCK F_CollectInput
  VAR_IN_OUT
      Data : ARRAY[1..50] OF BOOL;
  END_VAR
  VAR_INPUT
      TICK  : BOOL := 0;
      IN1   : BOOL := 0;
      IN2   : BOOL := 0;
      IN3   : BOOL := 0;
      IN4   : BOOL := 0;
      IN5   : BOOL := 0;
      RESET : BOOL := FALSE;
  END_VAR
  VAR_OUTPUT
      Finished : BOOL;
  END_VAR
  VAR
      j    : USINT := 1;
      tock : BOOL  := 0;
  END_VAR
  IF NOT RESET AND tock = NOT TICK THEN
      Data[j]   := IN1;
      Data[j+1] := IN2;
      Data[j+2] := IN3;
      Data[j+3] := IN4;
      Data[j+4] := IN5;
      j := j + 5;
      tock := TICK;
  ELSE
      j := 1;
      tock := 0;
  END_IF;
  Finished := (j > 50);
END_FUNCTION_BLOCK

PROGRAM Boiler
  VAR
    Data  : ARRAY[1..50] OF BOOL;
    Ready : BOOL;
    CollectInput : F_CollectInput;
  END_VAR
  VAR
    TICK     AT %IX1.0 : BOOL;
    IN1      AT %IX0.3 : BOOL;
    IN2      AT %IX0.4 : BOOL;
    IN3      AT %IX0.5 : BOOL;
    IN4      AT %IX0.6 : BOOL;
    IN5      AT %IX0.7 : BOOL;
    OutReady AT %QX0.0 : BOOL := FALSE;
    FeedNext AT %QX0.1 : BOOL := FALSE;
    Out      AT %QX0.2 : BOOL;
  END_VAR
  CollectInput(TICK:=TICK, IN1:=IN1, IN2:=IN2, IN3:=IN3, IN4:=IN4, IN5:=IN5);
  Ready := CollectInput.Finished;
  FeedNext := 1;
  IF Ready THEN
    Out := (NOT (NOT (Data[11] OR Data[43])));
    OutReady := 1;
    CollectInput(RESET:=TRUE);
  END_IF;
END_PROGRAM

CONFIGURATION Config0
  RESOURCE Res0 ON PLC
    TASK task0(INTERVAL := T#20ms,PRIORITY := 0);
    PROGRAM instance0 WITH task0 : Boiler;
  END_RESOURCE
END_CONFIGURATION

(* ---- RND-EXPR_monte-bucks-excon.st ---- *)
(*
This code implements a randomly grown symbolic expression:

IN34 & (((!(xor(xor(xor(xor(!(xor(xor(xor(xor(!(IN20), IN18), IN25), xor(xor(IN31 & IN24, IN21), !(IN25))), IN15)), !((xor(xor(IN46, IN23 | IN21), IN33 & IN48)) | (!(!(IN41))))), false | ((!(xor(xor(IN9, IN42), IN20))) & ((!(IN2)) | (IN13 | IN5)))), (IN5 | (xor(xor(xor(xor(xor(xor(IN50, false), IN48), !(IN16)), IN17 | IN4), IN27 & (IN16 | IN48)), (xor(xor(IN32, IN19), IN13)) & (IN3 | IN8)))) | (xor(xor(!((IN41 | IN14) & (!(IN7))), xor(xor(IN3, xor(xor(!(IN42), IN14), xor(xor(IN14, IN43), IN36))), xor(xor(IN39 & IN38, IN34 | IN41), IN9 & IN13))), !(!(!(IN28)))))), ((((xor(xor(false, IN39), IN18)) | (!(IN29))) & ((!(IN19)) & (!(IN13)))) | ((xor(xor(IN15, IN25 & IN5), false)) & ((xor(xor(IN32, IN20), IN50)) & (IN20 | IN41)))) | IN1))) | IN17) & (!(!(xor(xor((IN32 | (!(IN6 | (IN25 & IN4)))) & (((!(IN1)) & ((IN48 | IN37) | (!(IN28)))) | IN15), (!(xor(xor((IN13 | IN6) & (xor(xor(IN47, IN40), IN40)), IN17), IN5))) & ((xor(xor(!(IN7), xor(xor(IN50 & IN36, xor(xor(IN10, IN50), IN12)), IN4)), xor(xor(xor(xor(IN29, IN26), IN30), IN40 | IN2), xor(xor(IN27, IN25), IN42)))) & IN42)), IN16 | (!(xor(xor(!(IN16 | IN22), IN30), xor(xor(IN42 & IN47, IN40 | IN37), IN19 & IN32)))))))))

*)

FUNCTION_BLOCK F_CollectInput
  VAR_IN_OUT
      Data : ARRAY[1..50] OF BOOL;
  END_VAR
  VAR_INPUT
      TICK  : BOOL := 0;
      IN1   : BOOL := 0;
      IN2   : BOOL := 0;
      IN3   : BOOL := 0;
      IN4   : BOOL := 0;
      IN5   : BOOL := 0;
      RESET : BOOL := FALSE;
  END_VAR
  VAR_OUTPUT
      Finished : BOOL;
  END_VAR
  VAR
      j    : USINT := 1;
      tock : BOOL  := 0;
  END_VAR
  IF NOT RESET AND tock = NOT TICK THEN
      Data[j]   := IN1;
      Data[j+1] := IN2;
      Data[j+2] := IN3;
      Data[j+3] := IN4;
      Data[j+4] := IN5;
      j := j + 5;
      tock := TICK;
  ELSE
      j := 1;
      tock := 0;
  END_IF;
  Finished := (j > 50);
END_FUNCTION_BLOCK

PROGRAM Boiler
  VAR
    Data  : ARRAY[1..50] OF BOOL;
    Ready : BOOL;
    CollectInput : F_CollectInput;
  END_VAR
  VAR
    TICK     AT %IX1.0 : BOOL;
    IN1      AT %IX0.3 : BOOL;
    IN2      AT %IX0.4 : BOOL;
    IN3      AT %IX0.5 : BOOL;
    IN4      AT %IX0.6 : BOOL;
    IN5      AT %IX0.7 : BOOL;
    OutReady AT %QX0.0 : BOOL := FALSE;
    FeedNext AT %QX0.1 : BOOL := FALSE;
    Out      AT %QX0.2 : BOOL;
  END_VAR
  CollectInput(TICK:=TICK, IN1:=IN1, IN2:=IN2, IN3:=IN3, IN4:=IN4, IN5:=IN5);
  Ready := CollectInput.Finished;
  FeedNext := 1;
  IF Ready THEN
    Out := (Data[34] AND (((NOT (((((NOT (((((NOT Data[20]) XOR Data[18]) XOR Data[25]) XOR (((Data[31] AND Data[24]) XOR Data[21]) XOR (NOT Data[25]))) XOR Data[15])) XOR (NOT (((Data[46] XOR (Data[23] OR Data[21])) XOR (Data[33] AND Data[48])) OR (NOT (NOT Data[41]))))) XOR (FALSE OR ((NOT ((Data[9] XOR Data[42]) XOR Data[20])) AND ((NOT Data[2]) OR (Data[13] OR Data[5]))))) XOR ((Data[5] OR ((((((Data[50] XOR FALSE) XOR Data[48]) XOR (NOT Data[16])) XOR (Data[17] OR Data[4])) XOR (Data[27] AND (Data[16] OR Data[48]))) XOR (((Data[32] XOR Data[19]) XOR Data[13]) AND (Data[3] OR Data[8])))) OR (((NOT ((Data[41] OR Data[14]) AND (NOT Data[7]))) XOR ((Data[3] XOR (((NOT Data[42]) XOR Data[14]) XOR ((Data[14] XOR Data[43]) XOR Data[36]))) XOR (((Data[39] AND Data[38]) XOR (Data[34] OR Data[41])) XOR (Data[9] AND Data[13])))) XOR (NOT (NOT (NOT Data[28])))))) XOR ((((((FALSE XOR Data[39]) XOR Data[18]) OR (NOT Data[29])) AND ((NOT Data[19]) AND (NOT Data[13]))) OR (((Data[15] XOR (Data[25] AND Data[5])) XOR FALSE) AND (((Data[32] XOR Data[20]) XOR Data[50]) AND (Data[20] OR Data[41])))) OR Data[1]))) OR Data[17]) AND (NOT (NOT ((((Data[32] OR (NOT (Data[6] OR (Data[25] AND Data[4])))) AND (((NOT Data[1]) AND ((Data[48] OR Data[37]) OR (NOT Data[28]))) OR Data[15])) XOR ((NOT ((((Data[13] OR Data[6]) AND ((Data[47] XOR Data[40]) XOR Data[40])) XOR Data[17]) XOR Data[5])) AND ((((NOT Data[7]) XOR (((Data[50] AND Data[36]) XOR ((Data[10] XOR Data[50]) XOR Data[12])) XOR Data[4])) XOR ((((Data[29] XOR Data[26]) XOR Data[30]) XOR (Data[40] OR Data[2])) XOR ((Data[27] XOR Data[25]) XOR Data[42]))) AND Data[42]))) XOR (Data[16] OR (NOT (((NOT (Data[16] OR Data[22])) XOR Data[30]) XOR (((Data[42] AND Data[47]) XOR (Data[40] OR Data[37])) XOR (Data[19] AND Data[32]))))))))));
    OutReady := 1;
    CollectInput(RESET:=TRUE);
  END_IF;
END_PROGRAM

CONFIGURATION Config0
  RESOURCE Res0 ON PLC
    TASK task0(INTERVAL := T#20ms,PRIORITY := 0);
    PROGRAM instance0 WITH task0 : Boiler;
  END_RESOURCE
END_CONFIGURATION

(* ---- RND-EXPR_mopes-dicot-nixed.st ---- *)
(*
This code implements a randomly grown symbolic expression:

IN18 | (((xor(xor(xor(xor(IN17 | (xor(xor(IN20 | IN31, !((IN23 | IN3) | (!(IN14)))), xor(xor((!(IN35)) | (!(IN43)), IN8), !(IN28 | IN33)))), false), IN38 & IN24), ((IN39 | (((IN32 | true) | (!(IN47))) | ((xor(xor(IN25, IN42), IN28)) | (IN42 | IN24)))) & ((((xor(xor(IN38, IN18), IN2)) | (IN4 & IN11)) | ((!(IN45)) & (IN8 | IN28))) | (!((!(IN50)) & IN24)))) & (xor(xor(IN18, ((xor(xor(IN35 & IN33, false & IN2), !(IN32))) & (!(IN19 & IN38))) & ((!(xor(xor(IN7, IN2), IN18))) & ((xor(xor(IN48, IN26), false)) & (xor(xor(IN46, IN38), IN13))))), xor(xor(xor(xor(IN13 | (xor(xor(IN37, IN12), IN43)), IN36), xor(xor(IN17 | true, IN49), IN2)), (!(IN33 & IN19)) & IN43), IN7)))), xor(xor(xor(xor(xor(xor(((xor(xor(IN14, IN2), IN34)) & (xor(xor(IN43, IN41), IN11))) | ((IN34 & IN13) | (IN14 & IN33)), !(xor(xor(!(IN26), !(IN28)), !(IN43)))), (xor(xor(IN30, xor(xor(IN38, IN10), IN28)), xor(xor(IN36, IN49), IN11))) | IN9), xor(xor(xor(xor(!(xor(xor(IN48, IN48), IN47)), (!(IN23)) | (IN30 | IN42)), xor(xor(IN21 & IN37, IN19), IN31)), (!(IN28)) | IN38), xor(xor(IN31, !(!(IN19))), IN45))), (xor(xor(IN19, IN15), xor(xor(xor(xor(IN5, IN27), IN1), false), !(IN13)))) & (IN14 & (xor(xor(IN13 & IN11, IN1), xor(xor(true, IN33), IN46))))), IN37), IN6))) | (!(xor(xor((!(((IN13 | IN14) & IN11) | (xor(xor(IN46 & IN42, xor(xor(IN32, IN1), IN3)), !(IN7))))) & IN26, IN17 | IN13), (!(((!(IN34)) & (true & IN40)) & ((xor(xor(IN3, IN6), IN24)) & IN30))) & (((IN21 & (IN16 & IN37)) | (xor(xor(xor(xor(IN47, IN22), IN46), !(IN28)), IN6 | IN26))) | (((xor(xor(IN10, IN47), IN41)) & IN19) | ((!(IN12)) | (!(IN20))))))))) & IN32)

*)

FUNCTION_BLOCK F_CollectInput
  VAR_IN_OUT
      Data : ARRAY[1..50] OF BOOL;
  END_VAR
  VAR_INPUT
      TICK  : BOOL := 0;
      IN1   : BOOL := 0;
      IN2   : BOOL := 0;
      IN3   : BOOL := 0;
      IN4   : BOOL := 0;
      IN5   : BOOL := 0;
      RESET : BOOL := FALSE;
  END_VAR
  VAR_OUTPUT
      Finished : BOOL;
  END_VAR
  VAR
      j    : USINT := 1;
      tock : BOOL  := 0;
  END_VAR
  IF NOT RESET AND tock = NOT TICK THEN
      Data[j]   := IN1;
      Data[j+1] := IN2;
      Data[j+2] := IN3;
      Data[j+3] := IN4;
      Data[j+4] := IN5;
      j := j + 5;
      tock := TICK;
  ELSE
      j := 1;
      tock := 0;
  END_IF;
  Finished := (j > 50);
END_FUNCTION_BLOCK

PROGRAM Boiler
  VAR
    Data  : ARRAY[1..50] OF BOOL;
    Ready : BOOL;
    CollectInput : F_CollectInput;
  END_VAR
  VAR
    TICK     AT %IX1.0 : BOOL;
    IN1      AT %IX0.3 : BOOL;
    IN2      AT %IX0.4 : BOOL;
    IN3      AT %IX0.5 : BOOL;
    IN4      AT %IX0.6 : BOOL;
    IN5      AT %IX0.7 : BOOL;
    OutReady AT %QX0.0 : BOOL := FALSE;
    FeedNext AT %QX0.1 : BOOL := FALSE;
    Out      AT %QX0.2 : BOOL;
  END_VAR
  CollectInput(TICK:=TICK, IN1:=IN1, IN2:=IN2, IN3:=IN3, IN4:=IN4, IN5:=IN5);
  Ready := CollectInput.Finished;
  FeedNext := 1;
  IF Ready THEN
    Out := (Data[18] OR (((((((Data[17] OR (((Data[20] OR Data[31]) XOR (NOT ((Data[23] OR Data[3]) OR (NOT Data[14])))) XOR ((((NOT Data[35]) OR (NOT Data[43])) XOR Data[8]) XOR (NOT (Data[28] OR Data[33]))))) XOR FALSE) XOR (Data[38] AND Data[24])) XOR (((Data[39] OR (((Data[32] OR TRUE) OR (NOT Data[47])) OR (((Data[25] XOR Data[42]) XOR Data[28]) OR (Data[42] OR Data[24])))) AND (((((Data[38] XOR Data[18]) XOR Data[2]) OR (Data[4] AND Data[11])) OR ((NOT Data[45]) AND (Data[8] OR Data[28]))) OR (NOT ((NOT Data[50]) AND Data[24])))) AND ((Data[18] XOR (((((Data[35] AND Data[33]) XOR (FALSE AND Data[2])) XOR (NOT Data[32])) AND (NOT (Data[19] AND Data[38]))) AND ((NOT ((Data[7] XOR Data[2]) XOR Data[18])) AND (((Data[48] XOR Data[26]) XOR FALSE) AND ((Data[46] XOR Data[38]) XOR Data[13]))))) XOR (((((Data[13] OR ((Data[37] XOR Data[12]) XOR Data[43])) XOR Data[36]) XOR (((Data[17] OR TRUE) XOR Data[49]) XOR Data[2])) XOR ((NOT (Data[33] AND Data[19])) AND Data[43])) XOR Data[7])))) XOR ((((((((((Data[14] XOR Data[2]) XOR Data[34]) AND ((Data[43] XOR Data[41]) XOR Data[11])) OR ((Data[34] AND Data[13]) OR (Data[14] AND Data[33]))) XOR (NOT (((NOT Data[26]) XOR (NOT Data[28])) XOR (NOT Data[43])))) XOR (((Data[30] XOR ((Data[38] XOR Data[10]) XOR Data[28])) XOR ((Data[36] XOR Data[49]) XOR Data[11])) OR Data[9])) XOR (((((NOT ((Data[48] XOR Data[48]) XOR Data[47])) XOR ((NOT Data[23]) OR (Data[30] OR Data[42]))) XOR (((Data[21] AND Data[37]) XOR Data[19]) XOR Data[31])) XOR ((NOT Data[28]) OR Data[38])) XOR ((Data[31] XOR (NOT (NOT Data[19]))) XOR Data[45]))) XOR (((Data[19] XOR Data[15]) XOR ((((Data[5] XOR Data[27]) XOR Data[1]) XOR FALSE) XOR (NOT Data[13]))) AND (Data[14] AND (((Data[13] AND Data[11]) XOR Data[1]) XOR ((TRUE XOR Data[33]) XOR Data[46]))))) XOR Data[37]) XOR Data[6])) OR (NOT ((((NOT (((Data[13] OR Data[14]) AND Data[11]) OR (((Data[46] AND Data[42]) XOR ((Data[32] XOR Data[1]) XOR Data[3])) XOR (NOT Data[7])))) AND Data[26]) XOR (Data[17] OR Data[13])) XOR ((NOT (((NOT Data[34]) AND (TRUE AND Data[40])) AND (((Data[3] XOR Data[6]) XOR Data[24]) AND Data[30]))) AND (((Data[21] AND (Data[16] AND Data[37])) OR ((((Data[47] XOR Data[22]) XOR Data[46]) XOR (NOT Data[28])) XOR (Data[6] OR Data[26]))) OR ((((Data[10] XOR Data[47]) XOR Data[41]) AND Data[19]) OR ((NOT Data[12]) OR (NOT Data[20])))))))) AND Data[32]));
    OutReady := 1;
    CollectInput(RESET:=TRUE);
  END_IF;
END_PROGRAM

CONFIGURATION Config0
  RESOURCE Res0 ON PLC
    TASK task0(INTERVAL := T#20ms,PRIORITY := 0);
    PROGRAM instance0 WITH task0 : Boiler;
  END_RESOURCE
END_CONFIGURATION
